(* IEC 61131-3 sources: plc-st-coding-agent/progress/evidence/f14_v14_remaining_20261113/jobs/custom_minimax-m27 (part 7) *)

(* ---- self-hard-01.raw_candidate_02.st ---- *)
FUNCTION_BLOCK FB
VAR_INPUT
    flowLow   : BOOL;
    ackBtn    : BOOL;
    sensorOK  : BOOL;
END_VAR
VAR_OUTPUT
    alarmActive : BOOL;
    alarmAcked  : BOOL;
    highHigh    : BOOL;
END_VAR
VAR
    prev_flowLow  : BOOL := FALSE;
    prev_ackBtn   : BOOL := FALSE;
    prev_alarmActive : BOOL := FALSE;
    prev_alarmAcked  : BOOL := FALSE;
END_VAR
VAR_TEMP
    ackRising : BOOL;
END_VAR
(* ENGINEERING_CONTRACT
   ISA-18.2 four-state alarm (unack-active / unack-cleared / acked-active / acked-cleared):
   ┌──────────────────┬───────────────┬──────────────────────────────────────────────┐
   │ Output / State   │ Activation    │ Retention / Reset / Deactivation              │
   ├──────────────────┼───────────────┼──────────────────────────────────────────────┤
   │ alarmActive      │ flowLow rising│ Held until condition cleared AND alarmAcked   │
   │                  │ edge          │ (no self-clear without explicit ack)         │
   ├──────────────────┼───────────────┼──────────────────────────────────────────────┤
   │ alarmAcked       │ 1) ackBtn     │ Held across scans; reset only when acked-btn │
   │                  │    rising edge│    pressed while condition gone (clears both)│
   │                  │ 2) condition  │                                              │
   │                  │    cleared    │                                              │
   │                  │    (prev unack│                                              │
   │                  │    active)    │                                              │
   ├──────────────────┼───────────────┼──────────────────────────────────────────────┤
   │ highHigh         │ sensorOK=FALSE│ Auto-cleared when sensorOK returns TRUE      │
   │                  │ (same scan)   │ (independent, never inhibits low alarm)     │
   └──────────────────┴───────────────┴──────────────────────────────────────────────┘
   Boundaries:
     - alarmActive retained across scans when !alarmAcked (PUB001/PUB002/PUB005)
     - highHigh = NOT sensorOK  (PUB004/PUB016)
     - ackBtn rising-edge only; same-scan evaluation (PUB006/PUB007/PUB014)
     - No timers or hidden state; all VAR static (PUB008)
   Supported formal properties:
     [S1] G(flowLow & ackBtn -> alarmActive)
     [S2] G(alarmActive & !alarmAcked & X(flowLow) -> X(alarmActive))
     [S3] G(!sensorOK -> highHigh)
     [S4] G(rising(ackBtn) & flowLow -> alarmAcked)
     [S5] G(highHigh <-> !sensorOK)
     [S6] alarmActive FSM (see state table above)
     [S7] alarmAcked FSM (see state table above)
*)
    (* Rising-edge detection *)
    ackRising := ackBtn AND NOT prev_ackBtn;

    (* ── High-priority alarm: sensor wire-break ── *)
    highHigh := NOT sensorOK;  (* PUB004/PUB016, PUB034: auto-clear when OK *)

    (* ── Four-state low-priority alarm ── *)

    (* Condition gone transitions *)
    IF flowLow THEN
        (* Condition still present *)
        alarmActive := TRUE;
        IF ackRising THEN
            alarmAcked := TRUE;  (* acked while condition present: acked-active *)
        END_IF;
    ELSE
        (* Condition currently gone *)
        IF prev_flowLow THEN
            (* Just-cleared edge: alarm can't vanish unacknowledged *)
            IF alarmActive AND NOT alarmAcked THEN
                alarmAcked := TRUE;   (* unack-active → acked-cleared *)
            END_IF;
            (* acked-cleared stays active until user presses ack *)
            IF alarmActive AND alarmAcked THEN
                (* stay acked-cleared; handled below after ack check *)
            END_IF;
        END_IF;

        (* Transition out of acked-cleared on explicit acknowledge *)
        IF alarmActive AND alarmAcked AND ackRising THEN
            alarmActive := FALSE;
            alarmAcked  := FALSE;
        END_IF;

        (* No active alarm and not just cleared → cleared state *)
        IF NOT alarmActive THEN
            alarmAcked := FALSE;
        END_IF;
    END_IF;

    (* Persist alarmActive when condition present but not yet acked *)
    IF flowLow AND prev_flowLow AND alarmActive AND NOT alarmAcked THEN
        alarmActive := TRUE;   (* hold unack-active across scans *)
    END_IF;

    (* Shift-register for next scan *)
    prev_flowLow     := flowLow;
    prev_ackBtn      := ackBtn;
    prev_alarmActive := alarmActive;
    prev_alarmAcked  := alarmAcked;
END_FUNCTION_BLOCK

(* ---- self-hard-01.raw_candidate_03.st ---- *)
FUNCTION_BLOCK FB
VAR_INPUT
    flowLow   : BOOL;
    ackBtn    : BOOL;
    sensorOK  : BOOL;
END_VAR
VAR_OUTPUT
    alarmActive : BOOL;
    alarmAcked  : BOOL;
    highHigh    : BOOL;
END_VAR
VAR
    prev_flowLow  : BOOL := FALSE;
    prev_ackBtn   : BOOL := FALSE;
    prev_alarmActive : BOOL := FALSE;
    prev_alarmAcked  : BOOL := FALSE;
END_VAR
VAR_TEMP
    ackRising : BOOL;
END_VAR
(* ENGINEERING_CONTRACT
   ISA-18.2 four-state alarm (unack-active / unack-cleared / acked-active / acked-cleared):
   ┌──────────────────┬───────────────┬──────────────────────────────────────────────┐
   │ Output / State   │ Activation    │ Retention / Reset / Deactivation              │
   ├──────────────────┼───────────────┼──────────────────────────────────────────────┤
   │ alarmActive      │ flowLow rising│ Held until condition cleared AND alarmAcked   │
   │                  │ edge          │ (no self-clear without explicit ack)         │
   ├──────────────────┼───────────────┼──────────────────────────────────────────────┤
   │ alarmAcked       │ 1) ackBtn     │ Held across scans; reset only when acked-btn │
   │                  │    rising edge│    pressed while condition gone (clears both)│
   │                  │ 2) condition  │                                              │
   │                  │    cleared    │                                              │
   │                  │    (prev unack│                                              │
   │                  │    active)    │                                              │
   ├──────────────────┼───────────────┼──────────────────────────────────────────────┤
   │ highHigh         │ sensorOK=FALSE│ Auto-cleared when sensorOK returns TRUE      │
   │                  │ (same scan)   │ (independent, never inhibits low alarm)     │
   └──────────────────┴───────────────┴──────────────────────────────────────────────┘
   Boundaries:
     - alarmActive retained across scans when !alarmAcked (PUB001/PUB002/PUB005)
     - highHigh = NOT sensorOK  (PUB004/PUB016)
     - ackBtn rising-edge only; same-scan evaluation (PUB006/PUB007/PUB014)
     - No timers or hidden state; all VAR static (PUB008)
   Supported formal properties:
     [S1] G(flowLow & ackBtn -> alarmActive)
     [S2] G(alarmActive & !alarmAcked & X(flowLow) -> X(alarmActive))
     [S3] G(!sensorOK -> highHigh)
     [S4] G(rising(ackBtn) & flowLow -> alarmAcked)
     [S5] G(highHigh <-> !sensorOK)
     [S6] alarmActive FSM (see state table above)
     [S7] alarmAcked FSM (see state table above)
*)
    ackRising := ackBtn AND NOT prev_ackBtn;

    (* ── High-priority alarm: sensor wire-break ── *)
    highHigh := NOT sensorOK;  (* PUB004/PUB016, PUB034: auto-clear when OK *)

    (* ── Four-state low-priority alarm ── *)

    (* Condition gone transitions *)
    IF flowLow THEN
        (* Condition still present *)
        alarmActive := TRUE;
        IF ackRising THEN
            alarmAcked := TRUE;  (* acked while condition present: acked-active *)
        END_IF;
    ELSE
        (* Condition currently gone *)
        IF prev_flowLow THEN
            (* Just-cleared edge: alarm can't vanish unacknowledged *)
            IF alarmActive AND NOT alarmAcked THEN
                alarmAcked := TRUE;   (* unack-active → acked-cleared *)
            END_IF;
            (* acked-cleared stays active until user presses ack *)
            IF alarmActive AND alarmAcked THEN
                (* stay acked-cleared; handled below after ack check *)
            END_IF;
        END_IF;

        (* Transition out of acked-cleared on explicit acknowledge *)
        IF alarmActive AND alarmAcked AND ackRising THEN
            alarmActive := FALSE;
            alarmAcked  := FALSE;
        END_IF;

        (* No active alarm and not just cleared → cleared state *)
        IF NOT alarmActive THEN
            alarmAcked := FALSE;
        END_IF;
    END_IF;

    (* Persist alarmActive when condition present but not yet acked *)
    IF flowLow AND prev_flowLow AND alarmActive AND NOT alarmAcked THEN
        alarmActive := TRUE;   (* hold unack-active across scans *)
    END_IF;

    (* Shift-register for next scan *)
    prev_flowLow     := flowLow;
    prev_ackBtn      := ackBtn;
    prev_alarmActive := alarmActive;
    prev_alarmAcked  := alarmAcked;
END_FUNCTION_BLOCK

(* ---- self-hard-02.candidate_01.st ---- *)
FUNCTION_BLOCK FB
VAR_INPUT
    startBtn   : BOOL;
    abortBtn   : BOOL;
    setpoint   : REAL;
    pv         : REAL;
    maxDuration: INT;
END_VAR
VAR_OUTPUT
    elapsed : INT := 0;
    phase   : INT := 0;
    timeout : BOOL := FALSE;
END_VAR
VAR
    prev_startBtn : BOOL := FALSE;
    prev_abortBtn : BOOL := FALSE;
END_VAR

(* ENGINEERING_CONTRACT
  PUB001-003: Initial (phase,elapsed,timeout)=(0,0,FALSE) on cold-start.
  PUB004:    maxDuration is a positive integer scan-count threshold.
  PUB005-006: Priority order per scan: (1) abort, (2) new start rising edge,
              (3) running count. No external clock or TON used.
  PUB007:    abortBtn=TRUE  → phase=9 immediately; elapsed & timeout frozen.
             A consumed rising edge cannot re-trigger without a release-press.
  PUB008:    New start rising edge (no abort) → phase=1,elapsed=0,timeout=FALSE.
             Start scan does NOT increment elapsed.
  PUB009:    When prev phase∈{1,2}: elapsed += 1 first, then threshold check.
  PUB010:    If elapsed >= maxDuration → timeout=TRUE, phase=3 (takes priority
             over pv/setpoint check). Else if pv>=setpoint → phase=2, else phase=1.
  PUB011-012: phase=3 (complete) and phase=9 (aborted) freeze elapsed & timeout
              until a new valid start or abort event.
  S1-S5/N10-S1..S6: All formal properties encoded in conditional branches.
  Units: elapsed in scan-pairs; maxDuration in scan-pairs; no time dimension.
*)
(* CONTRACT_RULES
  []
*)

VAR
    tmp_risingStart : BOOL;
    tmp_risingAbort : BOOL;
    tmp_wasRunning  : BOOL;
    tmp_prevPhase   : INT;
    tmp_prevTimeout : BOOL;
END_VAR

tmp_risingStart := startBtn AND NOT prev_startBtn;
tmp_risingAbort := abortBtn  AND NOT prev_abortBtn;
tmp_prevPhase   := phase;
tmp_prevTimeout := timeout;

IF tmp_risingAbort THEN
    // PUB007: abort priority over same-scan rising start; freeze counters
    phase   := 9;
    // elapsed, timeout unchanged
ELSIF tmp_risingStart THEN
    // PUB008: new batch, start scan not counted
    phase    := 1;
    elapsed  := 0;
    timeout  := FALSE;
ELSIF (tmp_prevPhase = 1) OR (tmp_prevPhase = 2) THEN
    // PUB009: running phase → increment elapsed, then evaluate timeout/transition
    elapsed := elapsed + 1;
    IF elapsed >= maxDuration THEN
        // PUB010: timeout reached → complete; pv check skipped
        timeout := TRUE;
        phase   := 3;
    ELSIF pv >= setpoint THEN
        phase := 2;
    ELSE
        phase := 1;
    END_IF;
ELSIF (tmp_prevPhase = 3) OR (tmp_prevPhase = 9) THEN
    // PUB011-012: terminal states retain counters
    phase   := tmp_prevPhase;
    timeout := tmp_prevTimeout;
ELSE
    // idle (phase=0) with no start edge: hold state
    phase   := 0;
END_IF;

prev_startBtn := startBtn;
prev_abortBtn := abortBtn;
END_FUNCTION_BLOCK

(* ---- self-hard-02.patch_base_02.st ---- *)
FUNCTION_BLOCK FB
VAR_INPUT
    startBtn   : BOOL;
    abortBtn   : BOOL;
    setpoint   : REAL;
    pv         : REAL;
    maxDuration: INT;
END_VAR
VAR_OUTPUT
    elapsed : INT := 0;
    phase   : INT := 0;
    timeout : BOOL := FALSE;
END_VAR
VAR
    prev_startBtn : BOOL := FALSE;
    prev_abortBtn : BOOL := FALSE;
END_VAR

(* ENGINEERING_CONTRACT
  PUB001-003: Initial (phase,elapsed,timeout)=(0,0,FALSE) on cold-start.
  PUB004:    maxDuration is a positive integer scan-count threshold.
  PUB005-006: Priority order per scan: (1) abort, (2) new start rising edge,
              (3) running count. No external clock or TON used.
  PUB007:    abortBtn=TRUE  → phase=9 immediately; elapsed & timeout frozen.
             A consumed rising edge cannot re-trigger without a release-press.
  PUB008:    New start rising edge (no abort) → phase=1,elapsed=0,timeout=FALSE.
             Start scan does NOT increment elapsed.
  PUB009:    When prev phase∈{1,2}: elapsed += 1 first, then threshold check.
  PUB010:    If elapsed >= maxDuration → timeout=TRUE, phase=3 (takes priority
             over pv/setpoint check). Else if pv>=setpoint → phase=2, else phase=1.
  PUB011-012: phase=3 (complete) and phase=9 (aborted) freeze elapsed & timeout
              until a new valid start or abort event.
  S1-S5/N10-S1..S6: All formal properties encoded in conditional branches.
  Units: elapsed in scan-pairs; maxDuration in scan-pairs; no time dimension.
*)
(* CONTRACT_RULES
  []
*)

VAR
    tmp_risingStart : BOOL;
    tmp_risingAbort : BOOL;
    tmp_wasRunning  : BOOL;
    tmp_prevPhase   : INT;
    tmp_prevTimeout : BOOL;
END_VAR

tmp_risingStart := startBtn AND NOT prev_startBtn;
tmp_risingAbort := abortBtn  AND NOT prev_abortBtn;
tmp_prevPhase   := phase;
tmp_prevTimeout := timeout;

IF tmp_risingAbort THEN
    // PUB007: abort priority over same-scan rising start; freeze counters
    phase   := 9;
    // elapsed, timeout unchanged
ELSIF tmp_risingStart THEN
    // PUB008: new batch, start scan not counted
    phase    := 1;
    elapsed  := 0;
    timeout  := FALSE;
ELSIF (tmp_prevPhase = 1) OR (tmp_prevPhase = 2) THEN
    // PUB009: running phase → increment elapsed, then evaluate timeout/transition
    elapsed := elapsed + 1;
    IF elapsed >= maxDuration THEN
        // PUB010: timeout reached → complete; pv check skipped
        timeout := TRUE;
        phase   := 3;
    ELSIF pv >= setpoint THEN
        phase := 2;
    ELSE
        phase := 1;
    END_IF;
ELSIF (tmp_prevPhase = 3) OR (tmp_prevPhase = 9) THEN
    // PUB011-012: terminal states retain counters
    phase   := tmp_prevPhase;
    timeout := tmp_prevTimeout;
ELSE
    // idle (phase=0) with no start edge: hold state
    phase   := 0;
END_IF;

prev_startBtn := startBtn;
prev_abortBtn := abortBtn;
END_FUNCTION_BLOCK

(* ---- self-hard-02.patch_base_03.st ---- *)
FUNCTION_BLOCK FB
VAR_INPUT
    startBtn   : BOOL;
    abortBtn   : BOOL;
    setpoint   : REAL;
    pv         : REAL;
    maxDuration: INT;
END_VAR
VAR_OUTPUT
    elapsed : INT := 0;
    phase   : INT := 0;
    timeout : BOOL := FALSE;
END_VAR
VAR
    prev_startBtn : BOOL := FALSE;
    prev_abortBtn : BOOL := FALSE;
END_VAR

(* ENGINEERING_CONTRACT
  PUB001-003: Initial (phase,elapsed,timeout)=(0,0,FALSE) on cold-start.
  PUB004:    maxDuration is a positive integer scan-count threshold.
  PUB005-006: Priority order per scan: (1) abort, (2) new start rising edge,
              (3) running count. No external clock or TON used.
  PUB007:    abortBtn=TRUE  → phase=9 immediately; elapsed & timeout frozen.
             A consumed rising edge cannot re-trigger without a release-press.
  PUB008:    New start rising edge (no abort) → phase=1,elapsed=0,timeout=FALSE.
             Start scan does NOT increment elapsed.
  PUB009:    When prev phase∈{1,2}: elapsed += 1 first, then threshold check.
  PUB010:    If elapsed >= maxDuration → timeout=TRUE, phase=3 (takes priority
             over pv/setpoint check). Else if pv>=setpoint → phase=2, else phase=1.
  PUB011-012: phase=3 (complete) and phase=9 (aborted) freeze elapsed & timeout
              until a new valid start or abort event.
  S1-S5/N10-S1..S6: All formal properties encoded in conditional branches.
  Units: elapsed in scan-pairs; maxDuration in scan-pairs; no time dimension.
*)
(* CONTRACT_RULES
  []
*)

VAR
    tmp_risingStart : BOOL;
    tmp_risingAbort : BOOL;
    tmp_wasRunning  : BOOL;
    tmp_prevPhase   : INT;
    tmp_prevTimeout : BOOL;
END_VAR

tmp_risingStart := startBtn AND NOT prev_startBtn;
tmp_risingAbort := abortBtn  AND NOT prev_abortBtn;
tmp_prevPhase   := phase;
tmp_prevTimeout := timeout;

IF tmp_risingAbort THEN
    // PUB007: abort priority over same-scan rising start; freeze counters
    phase   := 9;
    // elapsed, timeout unchanged
ELSIF tmp_risingStart THEN
    // PUB008: new batch, start scan not counted
    phase    := 1;
    elapsed  := 0;
    timeout  := FALSE;
ELSIF (tmp_prevPhase = 1) OR (tmp_prevPhase = 2) THEN
    // PUB009: running phase → increment elapsed, then evaluate timeout/transition
    elapsed := elapsed + 1;
    IF elapsed >= maxDuration THEN
        // PUB010: timeout reached → complete; pv check skipped
        timeout := TRUE;
        phase   := 3;
    ELSIF pv >= setpoint THEN
        phase := 2;
    ELSE
        phase := 1;
    END_IF;
ELSIF (tmp_prevPhase = 3) OR (tmp_prevPhase = 9) THEN
    // PUB011-012: terminal states retain counters
    phase   := tmp_prevPhase;
    timeout := tmp_prevTimeout;
ELSE
    // idle (phase=0) with no start edge: hold state
    phase   := 0;
END_IF;

prev_startBtn := startBtn;
prev_abortBtn := abortBtn;
END_FUNCTION_BLOCK

(* ---- self-hard-02.raw_candidate_01.st ---- *)
FUNCTION_BLOCK FB
VAR_INPUT
    startBtn   : BOOL;
    abortBtn   : BOOL;
    setpoint   : REAL;
    pv         : REAL;
    maxDuration: INT;
END_VAR
VAR_OUTPUT
    elapsed : INT := 0;
    phase   : INT := 0;
    timeout : BOOL := FALSE;
END_VAR
VAR
    prev_startBtn : BOOL := FALSE;
    prev_abortBtn : BOOL := FALSE;
END_VAR

(* ENGINEERING_CONTRACT
  PUB001-003: Initial (phase,elapsed,timeout)=(0,0,FALSE) on cold-start.
  PUB004:    maxDuration is a positive integer scan-count threshold.
  PUB005-006: Priority order per scan: (1) abort, (2) new start rising edge,
              (3) running count. No external clock or TON used.
  PUB007:    abortBtn=TRUE  → phase=9 immediately; elapsed & timeout frozen.
             A consumed rising edge cannot re-trigger without a release-press.
  PUB008:    New start rising edge (no abort) → phase=1,elapsed=0,timeout=FALSE.
             Start scan does NOT increment elapsed.
  PUB009:    When prev phase∈{1,2}: elapsed += 1 first, then threshold check.
  PUB010:    If elapsed >= maxDuration → timeout=TRUE, phase=3 (takes priority
             over pv/setpoint check). Else if pv>=setpoint → phase=2, else phase=1.
  PUB011-012: phase=3 (complete) and phase=9 (aborted) freeze elapsed & timeout
              until a new valid start or abort event.
  S1-S5/N10-S1..S6: All formal properties encoded in conditional branches.
  Units: elapsed in scan-pairs; maxDuration in scan-pairs; no time dimension.
*)
(* CONTRACT_RULES
  []
*)

VAR
    tmp_risingStart : BOOL;
    tmp_risingAbort : BOOL;
    tmp_wasRunning  : BOOL;
    tmp_prevPhase   : INT;
    tmp_prevTimeout : BOOL;
END_VAR

tmp_risingStart := startBtn AND NOT prev_startBtn;
tmp_risingAbort := abortBtn  AND NOT prev_abortBtn;
tmp_prevPhase   := phase;
tmp_prevTimeout := timeout;

IF tmp_risingAbort THEN
    // PUB007: abort priority over same-scan rising start; freeze counters
    phase   := 9;
    // elapsed, timeout unchanged
ELSIF tmp_risingStart THEN
    // PUB008: new batch, start scan not counted
    phase    := 1;
    elapsed  := 0;
    timeout  := FALSE;
ELSIF (tmp_prevPhase = 1) OR (tmp_prevPhase = 2) THEN
    // PUB009: running phase → increment elapsed, then evaluate timeout/transition
    elapsed := elapsed + 1;
    IF elapsed >= maxDuration THEN
        // PUB010: timeout reached → complete; pv check skipped
        timeout := TRUE;
        phase   := 3;
    ELSIF pv >= setpoint THEN
        phase := 2;
    ELSE
        phase := 1;
    END_IF;
ELSIF (tmp_prevPhase = 3) OR (tmp_prevPhase = 9) THEN
    // PUB011-012: terminal states retain counters
    phase   := tmp_prevPhase;
    timeout := tmp_prevTimeout;
ELSE
    // idle (phase=0) with no start edge: hold state
    phase   := 0;
END_IF;

prev_startBtn := startBtn;
prev_abortBtn := abortBtn;
END_FUNCTION_BLOCK

(* ---- self-hard-03.candidate_01.st ---- *)
FUNCTION_BLOCK FB
VAR_INPUT
    pushEn  : BOOL;
    pushItem: INT;
    popEn   : BOOL;
END_VAR
VAR_IN_OUT
    fifo    : ARRAY[1..8] OF INT;
END_VAR
VAR_OUTPUT
    count   : INT := 0;
    full    : BOOL := FALSE;
    empty   : BOOL := TRUE;
    head    : INT := 0;
END_VAR
VAR
    pushR   : R_TRIG;
    popR    : R_TRIG;
    prevPushEn  : BOOL := FALSE;
    prevPopEn   : BOOL := FALSE;
    firstScan   : BOOL := TRUE;
END_VAR
VAR_TEMP
    prevCount   : INT;
END_VAR
END_VAR

(*
ENGINEERING_CONTRACT
================================================================================
PUB001 §rising-edge trigger·pushEn  → pushR.Q = pulse
PUB002 §rising-edge trigger·popEn   → popR.Q  = pulse
PUB003 §pop-first: popR then pushR; pop on count>0 only; push on count<8 only
PUB004 §output: count/empty/full/head consistent with array state each scan
PUB005 §fifo[1..count] compact, fifo[1]=head when count>0; others unspecified
PUB006 §full ∧ pushR only: count=8 (no change); empty ∧ popR only: count=0
PUB007 §simultaneous: prev(full)→pop frees slot, then push succeeds; count stays
PUB008 §simultaneous: prev(empty)→pop no-op, push succeeds; count = 1
PUB009 §head=0 when empty; head=fifo[1] when count>0
PUB010 §no hidden timers; state in VAR; edge detection via R_TRIG
PUB011 §IN_OUT fifo bound by caller; write to positions 1..count only
PUB012 §rising edge detected on transition FALSE→TRUE; hold does not repeat
PUB013 §shift-left only when count>1; count=1 pop leaves array unchanged
PUB014 §push to unfull queue: fifo[count]=pushItem on same scan
PUB015 §all outputs derived from same-scan state; no multi-scan buffering
PUB016 §R_TRIG/Q is valid only during the scan where rising edge occurs
PUB017 §first scan: init fifo to defined state via firstScan guard
PUB018 §prev(pushEn) tracked via prevPushEn; prev(popEn) via prevPopEn
PUB019 §S1: count∈[0,8], full↔count=8, empty↔count=0
PUB020 §S2: prev(full)∧pushR∧!popR → count=8
PUB021 §S3: prev(empty)∧popR∧!pushR → count=0
PUB022 §S6: count updated after pop+push chain; only successful actions change it
PUB023 §S7: accepted push → fifo[count]=pushItem
PUB024 §S8: shift-left by one position when pop succeeds; count>1 shift else nop
================================================================================
*)
BEGIN
    (* First-scan initialization: ensure defined state for fifo[1..8] *)
    IF firstScan THEN
        firstScan := FALSE;
        fifo[1] := 0;
        fifo[2] := 0;
        fifo[3] := 0;
        fifo[4] := 0;
        fifo[5] := 0;
        fifo[6] := 0;
        fifo[7] := 0;
        fifo[8] := 0;
    END_IF;

    (* Capture prevCount before any state mutation this scan *)
    prevCount := count;

    (* Detect rising edges per PUB001, PUB002, PUB012 *)
    pushR(CLK := pushEn);
    popR(CLK := popEn);

    (* PUB003 §pop-first order: handle pop before push *)
    IF popR.Q AND prevCount > 0 THEN
        (* S8 §shift-left only when count>1; count=1 pop leaves array unchanged (PUB013) *)
        IF prevCount > 1 THEN
            fifo[1] := fifo[2];
            fifo[2] := fifo[3];
            fifo[3] := fifo[4];
            fifo[4] := fifo[5];
            fifo[5] := fifo[6];
            fifo[6] := fifo[7];
            fifo[7] := fifo[8];
            fifo[8] := 0;
        ELSE
            (* count=1: array untouched, only count decrements (PUB013) *)
        END_IF;
        count := count - 1;
    END_IF;

    (* PUB003 §push on count<8; PUB007/PUB008 §simultaneous pop+push chain *)
    IF pushR.Q AND count < 8 THEN
        (* PUB014/PUB023 §accepted push: fifo[count]=pushItem (position BEFORE increment) *)
        fifo[count + 1] := pushItem;
        count := count + 1;
    END_IF;

    (* PUB004/PUB009 §derive output signals from final same-scan state *)
    full  := (count = 8);
    empty := (count = 0);
    IF count > 0 THEN
        head := fifo[1];
    ELSE
        head := 0;
    END_IF;

    (* Track previous input state for next-scan edge detection (PUB018) *)
    prevPushEn := pushEn;
    prevPopEn  := popEn;
END_FUNCTION_BLOCK

(* CONTRACT_RULES [] *)

(* ---- self-hard-03.candidate_02.st ---- *)
FUNCTION_BLOCK FB
VAR_INPUT
    pushEn  : BOOL;
    pushItem: INT;
    popEn   : BOOL;
END_VAR
VAR_IN_OUT
    fifo    : ARRAY[1..8] OF INT;
END_VAR
VAR_OUTPUT
    count   : INT := 0;
    full    : BOOL := FALSE;
    empty   : BOOL := TRUE;
    head    : INT := 0;
END_VAR
VAR
    pushR   : R_TRIG;
    popR    : R_TRIG;
    prevPushEn  : BOOL := FALSE;
    prevPopEn   : BOOL := FALSE;
    firstScan   : BOOL := TRUE;
END_VAR
VAR
    tmp_prevCount : INT;
END_VAR

(*
ENGINEERING_CONTRACT
================================================================================
PUB001 §rising-edge trigger·pushEn  → pushR.Q = pulse
PUB002 §rising-edge trigger·popEn   → popR.Q  = pulse
PUB003 §pop-first: popR then pushR; pop on count>0 only; push on count<8 only
PUB004 §output: count/empty/full/head consistent with array state each scan
PUB005 §fifo[1..count] compact, fifo[1]=head when count>0; others unspecified
PUB006 §full ∧ pushR only: count=8 (no change); empty ∧ popR only: count=0
PUB007 §simultaneous: prev(full)→pop frees slot, then push succeeds; count stays
PUB008 §simultaneous: prev(empty)→pop no-op, push succeeds; count = 1
PUB009 §head=0 when empty; head=fifo[1] when count>0
PUB010 §no hidden timers; state in VAR; edge detection via R_TRIG
PUB011 §IN_OUT fifo bound by caller; write to positions 1..count only
PUB012 §rising edge detected on transition FALSE→TRUE; hold does not repeat
PUB013 §shift-left only when count>1; count=1 pop leaves array unchanged
PUB014 §push to unfull queue: fifo[count]=pushItem on same scan
PUB015 §all outputs derived from same-scan state; no multi-scan buffering
PUB016 §R_TRIG/Q is valid only during the scan where rising edge occurs
PUB017 §first scan: init fifo to defined state via firstScan guard
PUB018 §prev(pushEn) tracked via prevPushEn; prev(popEn) via prevPopEn
PUB019 §S1: count∈[0,8], full↔count=8, empty↔count=0
PUB020 §S2: prev(full)∧pushR∧!popR → count=8
PUB021 §S3: prev(empty)∧popR∧!pushR → count=0
PUB022 §S6: count updated after pop+push chain; only successful actions change it
PUB023 §S7: accepted push → fifo[count]=pushItem
PUB024 §S8: shift-left by one position when pop succeeds; count>1 shift else nop
================================================================================
*)
    (* Capture tmp_prevCount before any state mutation this scan *)
    tmp_prevCount := count;

    (* Detect rising edges per PUB001, PUB002, PUB012 *)
    pushR(CLK := pushEn);
    popR(CLK := popEn);

    (* PUB003 §pop-first order: handle pop before push *)
    IF popR.Q AND tmp_prevCount > 0 THEN
        (* S8 §shift-left only when count>1; count=1 pop leaves array unchanged (PUB013) *)
        IF tmp_prevCount > 1 THEN
            fifo[1] := fifo[2];
            fifo[2] := fifo[3];
            fifo[3] := fifo[4];
            fifo[4] := fifo[5];
            fifo[5] := fifo[6];
            fifo[6] := fifo[7];
            fifo[7] := fifo[8];
            fifo[8] := 0;
        END_IF;
        count := count - 1;
    END_IF;

    (* PUB003 §push on count<8; PUB007/PUB008 §simultaneous pop+push chain *)
    IF pushR.Q AND count < 8 THEN
        (* PUB014/PUB023 §accepted push: fifo[count]=pushItem (position BEFORE increment) *)
        fifo[count + 1] := pushItem;
        count := count + 1;
    END_IF;

    (* PUB004/PUB009 §derive output signals from final same-scan state *)
    full  := (count = 8);
    empty := (count = 0);
    IF count > 0 THEN
        head := fifo[1];
    ELSE
        head := 0;
    END_IF;

    (* Track previous input state for next-scan edge detection (PUB018) *)
    prevPushEn := pushEn;
    prevPopEn  := popEn;
END_FUNCTION_BLOCK

(* CONTRACT_RULES [] *)

(* ---- self-hard-03.patch_base_02.st ---- *)
FUNCTION_BLOCK FB
VAR_INPUT
    pushEn  : BOOL;
    pushItem: INT;
    popEn   : BOOL;
END_VAR
VAR_IN_OUT
    fifo    : ARRAY[1..8] OF INT;
END_VAR
VAR_OUTPUT
    count   : INT := 0;
    full    : BOOL := FALSE;
    empty   : BOOL := TRUE;
    head    : INT := 0;
END_VAR
VAR
    pushR   : R_TRIG;
    popR    : R_TRIG;
    prevPushEn  : BOOL := FALSE;
    prevPopEn   : BOOL := FALSE;
    firstScan   : BOOL := TRUE;
END_VAR
VAR_TEMP
    prevCount   : INT;
END_VAR
END_VAR

(*
ENGINEERING_CONTRACT
================================================================================
PUB001 §rising-edge trigger·pushEn  → pushR.Q = pulse
PUB002 §rising-edge trigger·popEn   → popR.Q  = pulse
PUB003 §pop-first: popR then pushR; pop on count>0 only; push on count<8 only
PUB004 §output: count/empty/full/head consistent with array state each scan
PUB005 §fifo[1..count] compact, fifo[1]=head when count>0; others unspecified
PUB006 §full ∧ pushR only: count=8 (no change); empty ∧ popR only: count=0
PUB007 §simultaneous: prev(full)→pop frees slot, then push succeeds; count stays
PUB008 §simultaneous: prev(empty)→pop no-op, push succeeds; count = 1
PUB009 §head=0 when empty; head=fifo[1] when count>0
PUB010 §no hidden timers; state in VAR; edge detection via R_TRIG
PUB011 §IN_OUT fifo bound by caller; write to positions 1..count only
PUB012 §rising edge detected on transition FALSE→TRUE; hold does not repeat
PUB013 §shift-left only when count>1; count=1 pop leaves array unchanged
PUB014 §push to unfull queue: fifo[count]=pushItem on same scan
PUB015 §all outputs derived from same-scan state; no multi-scan buffering
PUB016 §R_TRIG/Q is valid only during the scan where rising edge occurs
PUB017 §first scan: init fifo to defined state via firstScan guard
PUB018 §prev(pushEn) tracked via prevPushEn; prev(popEn) via prevPopEn
PUB019 §S1: count∈[0,8], full↔count=8, empty↔count=0
PUB020 §S2: prev(full)∧pushR∧!popR → count=8
PUB021 §S3: prev(empty)∧popR∧!pushR → count=0
PUB022 §S6: count updated after pop+push chain; only successful actions change it
PUB023 §S7: accepted push → fifo[count]=pushItem
PUB024 §S8: shift-left by one position when pop succeeds; count>1 shift else nop
================================================================================
*)
BEGIN
    (* First-scan initialization: ensure defined state for fifo[1..8] *)
    IF firstScan THEN
        firstScan := FALSE;
        fifo[1] := 0;
        fifo[2] := 0;
        fifo[3] := 0;
        fifo[4] := 0;
        fifo[5] := 0;
        fifo[6] := 0;
        fifo[7] := 0;
        fifo[8] := 0;
    END_IF;

    (* Capture prevCount before any state mutation this scan *)
    prevCount := count;

    (* Detect rising edges per PUB001, PUB002, PUB012 *)
    pushR(CLK := pushEn);
    popR(CLK := popEn);

    (* PUB003 §pop-first order: handle pop before push *)
    IF popR.Q AND prevCount > 0 THEN
        (* S8 §shift-left only when count>1; count=1 pop leaves array unchanged (PUB013) *)
        IF prevCount > 1 THEN
            fifo[1] := fifo[2];
            fifo[2] := fifo[3];
            fifo[3] := fifo[4];
            fifo[4] := fifo[5];
            fifo[5] := fifo[6];
            fifo[6] := fifo[7];
            fifo[7] := fifo[8];
            fifo[8] := 0;
        ELSE
            (* count=1: array untouched, only count decrements (PUB013) *)
        END_IF;
        count := count - 1;
    END_IF;

    (* PUB003 §push on count<8; PUB007/PUB008 §simultaneous pop+push chain *)
    IF pushR.Q AND count < 8 THEN
        (* PUB014/PUB023 §accepted push: fifo[count]=pushItem (position BEFORE increment) *)
        fifo[count + 1] := pushItem;
        count := count + 1;
    END_IF;

    (* PUB004/PUB009 §derive output signals from final same-scan state *)
    full  := (count = 8);
    empty := (count = 0);
    IF count > 0 THEN
        head := fifo[1];
    ELSE
        head := 0;
    END_IF;

    (* Track previous input state for next-scan edge detection (PUB018) *)
    prevPushEn := pushEn;
    prevPopEn  := popEn;
END_FUNCTION_BLOCK

(* CONTRACT_RULES [] *)

(* ---- self-hard-03.raw_candidate_01.st ---- *)
FUNCTION_BLOCK FB
VAR_INPUT
    pushEn  : BOOL;
    pushItem: INT;
    popEn   : BOOL;
END_VAR
VAR_IN_OUT
    fifo    : ARRAY[1..8] OF INT;
END_VAR
VAR_OUTPUT
    count   : INT := 0;
    full    : BOOL := FALSE;
    empty   : BOOL := TRUE;
    head    : INT := 0;
END_VAR
VAR
    pushR   : R_TRIG;
    popR    : R_TRIG;
    prevPushEn  : BOOL := FALSE;
    prevPopEn   : BOOL := FALSE;
    firstScan   : BOOL := TRUE;
END_VAR
VAR_TEMP
    prevCount   : INT;
END_VAR
END_VAR

(*
ENGINEERING_CONTRACT
================================================================================
PUB001 §rising-edge trigger·pushEn  → pushR.Q = pulse
PUB002 §rising-edge trigger·popEn   → popR.Q  = pulse
PUB003 §pop-first: popR then pushR; pop on count>0 only; push on count<8 only
PUB004 §output: count/empty/full/head consistent with array state each scan
PUB005 §fifo[1..count] compact, fifo[1]=head when count>0; others unspecified
PUB006 §full ∧ pushR only: count=8 (no change); empty ∧ popR only: count=0
PUB007 §simultaneous: prev(full)→pop frees slot, then push succeeds; count stays
PUB008 §simultaneous: prev(empty)→pop no-op, push succeeds; count = 1
PUB009 §head=0 when empty; head=fifo[1] when count>0
PUB010 §no hidden timers; state in VAR; edge detection via R_TRIG
PUB011 §IN_OUT fifo bound by caller; write to positions 1..count only
PUB012 §rising edge detected on transition FALSE→TRUE; hold does not repeat
PUB013 §shift-left only when count>1; count=1 pop leaves array unchanged
PUB014 §push to unfull queue: fifo[count]=pushItem on same scan
PUB015 §all outputs derived from same-scan state; no multi-scan buffering
PUB016 §R_TRIG/Q is valid only during the scan where rising edge occurs
PUB017 §first scan: init fifo to defined state via firstScan guard
PUB018 §prev(pushEn) tracked via prevPushEn; prev(popEn) via prevPopEn
PUB019 §S1: count∈[0,8], full↔count=8, empty↔count=0
PUB020 §S2: prev(full)∧pushR∧!popR → count=8
PUB021 §S3: prev(empty)∧popR∧!pushR → count=0
PUB022 §S6: count updated after pop+push chain; only successful actions change it
PUB023 §S7: accepted push → fifo[count]=pushItem
PUB024 §S8: shift-left by one position when pop succeeds; count>1 shift else nop
================================================================================
*)
BEGIN
    (* First-scan initialization: ensure defined state for fifo[1..8] *)
    IF firstScan THEN
        firstScan := FALSE;
        fifo[1] := 0;
        fifo[2] := 0;
        fifo[3] := 0;
        fifo[4] := 0;
        fifo[5] := 0;
        fifo[6] := 0;
        fifo[7] := 0;
        fifo[8] := 0;
    END_IF

    (* Capture prevCount before any state mutation this scan *)
    prevCount := count;

    (* Detect rising edges per PUB001, PUB002, PUB012 *)
    pushR(CLK := pushEn);
    popR(CLK := popEn);

    (* PUB003 §pop-first order: handle pop before push *)
    IF popR.Q AND prevCount > 0 THEN
        (* S8 §shift-left only when count>1; count=1 pop leaves array unchanged (PUB013) *)
        IF prevCount > 1 THEN
            fifo[1] := fifo[2];
            fifo[2] := fifo[3];
            fifo[3] := fifo[4];
            fifo[4] := fifo[5];
            fifo[5] := fifo[6];
            fifo[6] := fifo[7];
            fifo[7] := fifo[8];
            fifo[8] := 0;
        ELSE
            (* count=1: array untouched, only count decrements (PUB013) *)
        END_IF
        count := count - 1;
    END_IF

    (* PUB003 §push on count<8; PUB007/PUB008 §simultaneous pop+push chain *)
    IF pushR.Q AND count < 8 THEN
        (* PUB014/PUB023 §accepted push: fifo[count]=pushItem (position BEFORE increment) *)
        fifo[count + 1] := pushItem;
        count := count + 1;
    END_IF

    (* PUB004/PUB009 §derive output signals from final same-scan state *)
    full  := (count = 8);
    empty := (count = 0);
    IF count > 0 THEN
        head := fifo[1];
    ELSE
        head := 0;
    END_IF

    (* Track previous input state for next-scan edge detection (PUB018) *)
    prevPushEn := pushEn;
    prevPopEn  := popEn;
END_FUNCTION_BLOCK

(* CONTRACT_RULES [] *)

(* ---- self-hard-03.raw_candidate_02.st ---- *)
FUNCTION_BLOCK FB
VAR_INPUT
    pushEn  : BOOL;
    pushItem: INT;
    popEn   : BOOL;
END_VAR
VAR_IN_OUT
    fifo    : ARRAY[1..8] OF INT;
END_VAR
VAR_OUTPUT
    count   : INT := 0;
    full    : BOOL := FALSE;
    empty   : BOOL := TRUE;
    head    : INT := 0;
END_VAR
VAR
    pushR   : R_TRIG;
    popR    : R_TRIG;
    prevPushEn  : BOOL := FALSE;
    prevPopEn   : BOOL := FALSE;
    firstScan   : BOOL := TRUE;
END_VAR
VAR
    tmp_prevCount : INT;
END_VAR

(*
ENGINEERING_CONTRACT
================================================================================
PUB001 §rising-edge trigger·pushEn  → pushR.Q = pulse
PUB002 §rising-edge trigger·popEn   → popR.Q  = pulse
PUB003 §pop-first: popR then pushR; pop on count>0 only; push on count<8 only
PUB004 §output: count/empty/full/head consistent with array state each scan
PUB005 §fifo[1..count] compact, fifo[1]=head when count>0; others unspecified
PUB006 §full ∧ pushR only: count=8 (no change); empty ∧ popR only: count=0
PUB007 §simultaneous: prev(full)→pop frees slot, then push succeeds; count stays
PUB008 §simultaneous: prev(empty)→pop no-op, push succeeds; count = 1
PUB009 §head=0 when empty; head=fifo[1] when count>0
PUB010 §no hidden timers; state in VAR; edge detection via R_TRIG
PUB011 §IN_OUT fifo bound by caller; write to positions 1..count only
PUB012 §rising edge detected on transition FALSE→TRUE; hold does not repeat
PUB013 §shift-left only when count>1; count=1 pop leaves array unchanged
PUB014 §push to unfull queue: fifo[count]=pushItem on same scan
PUB015 §all outputs derived from same-scan state; no multi-scan buffering
PUB016 §R_TRIG/Q is valid only during the scan where rising edge occurs
PUB017 §first scan: init fifo to defined state via firstScan guard
PUB018 §prev(pushEn) tracked via prevPushEn; prev(popEn) via prevPopEn
PUB019 §S1: count∈[0,8], full↔count=8, empty↔count=0
PUB020 §S2: prev(full)∧pushR∧!popR → count=8
PUB021 §S3: prev(empty)∧popR∧!pushR → count=0
PUB022 §S6: count updated after pop+push chain; only successful actions change it
PUB023 §S7: accepted push → fifo[count]=pushItem
PUB024 §S8: shift-left by one position when pop succeeds; count>1 shift else nop
================================================================================
*)
    (* Capture tmp_prevCount before any state mutation this scan *)
    tmp_prevCount := count;

    (* Detect rising edges per PUB001, PUB002, PUB012 *)
    pushR(CLK := pushEn);
    popR(CLK := popEn);

    (* PUB003 §pop-first order: handle pop before push *)
    IF popR.Q AND tmp_prevCount > 0 THEN
        (* S8 §shift-left only when count>1; count=1 pop leaves array unchanged (PUB013) *)
        IF tmp_prevCount > 1 THEN
            fifo[1] := fifo[2];
            fifo[2] := fifo[3];
            fifo[3] := fifo[4];
            fifo[4] := fifo[5];
            fifo[5] := fifo[6];
            fifo[6] := fifo[7];
            fifo[7] := fifo[8];
            fifo[8] := 0;
        END_IF;
        count := count - 1;
    END_IF;

    (* PUB003 §push on count<8; PUB007/PUB008 §simultaneous pop+push chain *)
    IF pushR.Q AND count < 8 THEN
        (* PUB014/PUB023 §accepted push: fifo[count]=pushItem (position BEFORE increment) *)
        fifo[count + 1] := pushItem;
        count := count + 1;
    END_IF;

    (* PUB004/PUB009 §derive output signals from final same-scan state *)
    full  := (count = 8);
    empty := (count = 0);
    IF count > 0 THEN
        head := fifo[1];
    ELSE
        head := 0;
    END_IF;

    (* Track previous input state for next-scan edge detection (PUB018) *)
    prevPushEn := pushEn;
    prevPopEn  := popEn;
END_FUNCTION_BLOCK

(* CONTRACT_RULES [] *)

(* ---- self-hard-04.candidate_01.st ---- *)
FUNCTION_BLOCK FB
VAR_INPUT
    demand     : INT;
    runHours   : ARRAY[1..5] OF LINT;
    rotated    : BOOL;
END_VAR
VAR_OUTPUT
    leadPump    : INT := 0;
    lagPump     : INT := 0;
    runningCount: INT := 0;
END_VAR
VAR
    prevDemand   : INT := 0;
    prevLeadPump : INT := 0;
    tmp_minHours : LINT;
    tmp_minPump  : INT;
    tmp_lagPump  : INT;
    tmp_lagHours : LINT;
    tmp_lagChanged: BOOL;
    i            : INT;
    clippedDemand: INT;
    demandIncrease: BOOL;
END_VAR
VAR_TEMP
    tmp_leadHours: LINT;
    tmp_leadPump : INT;
END_VAR
// ---------------------------------------------------------------------
// ENGINEERING_CONTRACT
// PubRefs: PUB001–PUB046
// State retention: leadPump/lagPump held across scans until demand=0 (PUB003/PUB004/PUB026)
//   or until hysteresis rotation condition satisfied (PUB009/PUB030)
// Output retention: runningCount strictly tracks clipped demand every scan (PUB001/PUB003)
//   lagPump retained when no trigger event occurs (PUB008/PUB042)
// Reset on demand=0: leadPump=lagPump=0 immediately this scan (PUB003/PUB027)
// Initial state (first scan): leadPump=0, lagPump=0, runningCount=0 (PUB029)
// Hysteresis: rotation only when runHours[prevLead] - min(runHours[*]) > 50 strictly (PUB030/PUB040)
// Lag trigger: initial selection OR lead change OR runningCount increase (PUB008/PUB043)
// Lag exclusion: leadPump never equals lagPump when demand>=2 (PUB003/PUB004)
// ---------------------------------------------------------------------
// CONTRACT_RULES
// (No unconditional Boolean output latches specified in this task)
// []

// Clip demand to 0..5
IF demand < 0 THEN
    clippedDemand := 0;
ELSIF demand > 5 THEN
    clippedDemand := 5;
ELSE
    clippedDemand := demand;
END_IF;

runningCount := clippedDemand;
demandIncrease := (clippedDemand > prevDemand);

// Compute global minimum (runHours, pump#) for hysteresis check
tmp_minHours := runHours[1];
tmp_minPump := 1;
FOR i := 2 TO 5 DO
    IF runHours[i] < tmp_minHours OR (runHours[i] = tmp_minHours AND i < tmp_minPump) THEN
        tmp_minHours := runHours[i];
        tmp_minPump := i;
    END_IF;
END_FOR;

// Demand zero: clear both outputs immediately
IF clippedDemand = 0 THEN
    leadPump := 0;
    lagPump := 0;
ELSE
    // Positive demand branch
    IF prevLeadPump = 0 THEN
        // PUB003/PUB026: Initial selection - pick (runHours, pump#) minimum as lead
        tmp_leadHours := runHours[1];
        tmp_leadPump := 1;
        FOR i := 2 TO 5 DO
            IF runHours[i] < tmp_leadHours OR (runHours[i] = tmp_leadHours AND i < tmp_leadPump) THEN
                tmp_leadHours := runHours[i];
                tmp_leadPump := i;
            END_IF;
        END_FOR;
        leadPump := tmp_leadPump;
        tmp_lagChanged := TRUE;
    ELSE
        // PUB009/PUB030: Subsequent scan - apply hysteresis rotation
        // Only switch if rotated=TRUE AND (prevLead runHours - min runHours) > 50 strictly
        IF rotated AND (runHours[prevLeadPump] - tmp_minHours > 50) THEN
            leadPump := tmp_minPump;
            tmp_lagChanged := TRUE;
        ELSE
            // PUB006/PUB042: No rotation request or hysteresis not met - retain lead
            leadPump := prevLeadPump;
            tmp_lagChanged := FALSE;
        END_IF;
    END_IF;

    // PUB008/PUB043: Lag pump selection (triggered by initial/lead-change/runningCount-increase)
    IF clippedDemand >= 2 THEN
        IF tmp_lagChanged OR demandIncrease THEN
            tmp_lagPump := 0;
            tmp_lagHours := LINT#16#7FFFFFFFFFFFFFFF;
            FOR i := 1 TO 5 DO
                IF i <> leadPump THEN
                    IF runHours[i] < tmp_lagHours OR (runHours[i] = tmp_lagHours AND i < tmp_lagPump) THEN
                        tmp_lagHours := runHours[i];
                        tmp_lagPump := i;
                    END_IF;
                END_IF;
            END_FOR;
            lagPump := tmp_lagPump;
        END_IF;
        // ELSE: retain prev lagPump (no assignment)
    ELSE
        // PUB003: demand = 1, lagPump must be 0
        lagPump := 0;
    END_IF;
END_IF;

// Update previous-state trackers for next scan
prevDemand := clippedDemand;
prevLeadPump := leadPump;
END_FUNCTION_BLOCK

(* ---- self-hard-04.raw_candidate_01.st ---- *)
FUNCTION_BLOCK FB
VAR_INPUT
    demand     : INT;
    runHours   : ARRAY[1..5] OF LINT;
    rotated    : BOOL;
END_VAR
VAR_OUTPUT
    leadPump    : INT := 0;
    lagPump     : INT := 0;
    runningCount: INT := 0;
END_VAR
VAR
    prevDemand   : INT := 0;
    prevLeadPump : INT := 0;
    tmp_minHours : LINT;
    tmp_minPump  : INT;
    tmp_lagPump  : INT;
    tmp_lagHours : LINT;
    tmp_lagChanged: BOOL;
    i            : INT;
    clippedDemand: INT;
    demandIncrease: BOOL;
END_VAR
VAR_TEMP
    tmp_leadHours: LINT;
    tmp_leadPump : INT;
END_VAR
// ---------------------------------------------------------------------
// ENGINEERING_CONTRACT
// PubRefs: PUB001–PUB046
// State retention: leadPump/lagPump held across scans until demand=0 (PUB003/PUB004/PUB026)
//   or until hysteresis rotation condition satisfied (PUB009/PUB030)
// Output retention: runningCount strictly tracks clipped demand every scan (PUB001/PUB003)
//   lagPump retained when no trigger event occurs (PUB008/PUB042)
// Reset on demand=0: leadPump=lagPump=0 immediately this scan (PUB003/PUB027)
// Initial state (first scan): leadPump=0, lagPump=0, runningCount=0 (PUB029)
// Hysteresis: rotation only when runHours[prevLead] - min(runHours[*]) > 50 strictly (PUB030/PUB040)
// Lag trigger: initial selection OR lead change OR runningCount increase (PUB008/PUB043)
// Lag exclusion: leadPump never equals lagPump when demand>=2 (PUB003/PUB004)
// ---------------------------------------------------------------------
// CONTRACT_RULES
// (No unconditional Boolean output latches specified in this task)
// []

// Clip demand to 0..5
IF demand < 0 THEN
    clippedDemand := 0;
ELSIF demand > 5 THEN
    clippedDemand := 5;
ELSE
    clippedDemand := demand;
END_IF

runningCount := clippedDemand;
demandIncrease := (clippedDemand > prevDemand);

// Compute global minimum (runHours, pump#) for hysteresis check
tmp_minHours := runHours[1];
tmp_minPump := 1;
FOR i := 2 TO 5 DO
    IF runHours[i] < tmp_minHours OR (runHours[i] = tmp_minHours AND i < tmp_minPump) THEN
        tmp_minHours := runHours[i];
        tmp_minPump := i;
    END_IF
END_FOR

// Demand zero: clear both outputs immediately
IF clippedDemand = 0 THEN
    leadPump := 0;
    lagPump := 0;
ELSE
    // Positive demand branch
    IF prevLeadPump = 0 THEN
        // PUB003/PUB026: Initial selection - pick (runHours, pump#) minimum as lead
        tmp_leadHours := runHours[1];
        tmp_leadPump := 1;
        FOR i := 2 TO 5 DO
            IF runHours[i] < tmp_leadHours OR (runHours[i] = tmp_leadHours AND i < tmp_leadPump) THEN
                tmp_leadHours := runHours[i];
                tmp_leadPump := i;
            END_IF
        END_FOR
        leadPump := tmp_leadPump;
        tmp_lagChanged := TRUE;
    ELSE
        // PUB009/PUB030: Subsequent scan - apply hysteresis rotation
        // Only switch if rotated=TRUE AND (prevLead runHours - min runHours) > 50 strictly
        IF rotated AND (runHours[prevLeadPump] - tmp_minHours > 50) THEN
            leadPump := tmp_minPump;
            tmp_lagChanged := TRUE;
        ELSE
            // PUB006/PUB042: No rotation request or hysteresis not met - retain lead
            leadPump := prevLeadPump;
            tmp_lagChanged := FALSE;
        END_IF
    END_IF

    // PUB008/PUB043: Lag pump selection (triggered by initial/lead-change/runningCount-increase)
    IF clippedDemand >= 2 THEN
        IF tmp_lagChanged OR demandIncrease THEN
            tmp_lagPump := 0;
            tmp_lagHours := LINT#16#7FFFFFFFFFFFFFFF;
            FOR i := 1 TO 5 DO
                IF i <> leadPump THEN
                    IF runHours[i] < tmp_lagHours OR (runHours[i] = tmp_lagHours AND i < tmp_lagPump) THEN
                        tmp_lagHours := runHours[i];
                        tmp_lagPump := i;
                    END_IF
                END_IF
            END_FOR
            lagPump := tmp_lagPump;
        END_IF
        // ELSE: retain prev lagPump (no assignment)
    ELSE
        // PUB003: demand = 1, lagPump must be 0
        lagPump := 0;
    END_IF
END_IF

// Update previous-state trackers for next scan
prevDemand := clippedDemand;
prevLeadPump := leadPump;
END_FUNCTION_BLOCK

(* ---- self-hard-05.candidate_01.st ---- *)
(* ENGINEERING_CONTRACT
1. tripLatched: activation is runRequest AND NOT flameOK; the trip is set in the same scan (PUB001, PUB003, PUB031).
2. tripLatched retention: remains TRUE until a rising resetBtn edge while runRequest=FALSE AND flameOK=FALSE (PUB002, PUB005, PUB032).
3. Reset priority: the safety-state rising edge clears an existing trip; an invalid reset edge has no effect (PUB032).
4. fuelPermit: combinational from runRequest, flameOK, and NOT tripLatched; no fuel is permitted while tripped (PUB003, PUB004, PUB007).
5. trimEnable/airTrim: active only with fuelPermit and no analyzer fault; trim is clamped to [-10,+10] (PUB009, PUB010, PUB011).
6. o2Fault: combinational analyzer validity/range fault; it removes trim only and never removes fuelPermit (PUB008, PUB012).
7. airCommand: fuelPermit permits the command; otherwise it is 0.0; permitted values are clamped to [0,100] (PUB006, PUB013, PUB014).
8. All outputs are sampled at scan end; no startup, purge, ignition, or BMS sequencing is included (PUB015).
9. Units: o2PV and air values are percent; airTrim limits are output bounds, not guaranteed reachable trim values.
10. Unspecified startup sequencing and external baseAir validity are not added as interlocks.
*)
(* CONTRACT_RULES [] *)

FUNCTION_BLOCK FB
VAR_INPUT
    runRequest : BOOL;
    flameOK : BOOL;
    o2Valid : BOOL;
    o2PV : REAL;
    baseAir : REAL;
    resetBtn : BOOL;
END_VAR

VAR_OUTPUT
    fuelPermit : BOOL;
    trimEnable : BOOL;
    airTrim : REAL;
    airCommand : REAL;
    tripLatched : BOOL;
    o2Fault : BOOL;
END_VAR

VAR
    tmp_resetPrev : BOOL := FALSE;
    tmp_resetRising : BOOL;
    tmp_rawTrim : REAL;
    tmp_rawCommand : REAL;
END_VAR

tmp_resetRising := resetBtn AND NOT tmp_resetPrev;

IF runRequest AND NOT flameOK THEN
    tripLatched := TRUE;
ELSIF tripLatched AND tmp_resetRising AND NOT runRequest AND NOT flameOK THEN
    tripLatched := FALSE;
END_IF;

tmp_resetPrev := resetBtn;

fuelPermit := runRequest AND flameOK AND NOT tripLatched;

o2Fault := NOT o2Valid OR o2PV < 0.0 OR o2PV > 21.0;
trimEnable := fuelPermit AND NOT o2Fault;

IF trimEnable THEN
    tmp_rawTrim := 2.0 * (2.0 - o2PV);
    IF tmp_rawTrim > 10.0 THEN
        airTrim := 10.0;
    ELSIF tmp_rawTrim < -10.0 THEN
        airTrim := -10.0;
    ELSE
        airTrim := tmp_rawTrim;
    END_IF;
ELSE
    airTrim := 0.0;
END_IF;

IF fuelPermit THEN
    tmp_rawCommand := baseAir + airTrim;
    IF tmp_rawCommand > 100.0 THEN
        airCommand := 100.0;
    ELSIF tmp_rawCommand < 0.0 THEN
        airCommand := 0.0;
    ELSE
        airCommand := tmp_rawCommand;
    END_IF;
ELSE
    airCommand := 0.0;
END_IF;

END_FUNCTION_BLOCK

(* ---- self-hard-05.raw_candidate_01.st ---- *)
(* ENGINEERING_CONTRACT
1. tripLatched: activation is runRequest AND NOT flameOK; the trip is set in the same scan (PUB001, PUB003, PUB031).
2. tripLatched retention: remains TRUE until a rising resetBtn edge while runRequest=FALSE AND flameOK=FALSE (PUB002, PUB005, PUB032).
3. Reset priority: the safety-state rising edge clears an existing trip; an invalid reset edge has no effect (PUB032).
4. fuelPermit: combinational from runRequest, flameOK, and NOT tripLatched; no fuel is permitted while tripped (PUB003, PUB004, PUB007).
5. trimEnable/airTrim: active only with fuelPermit and no analyzer fault; trim is clamped to [-10,+10] (PUB009, PUB010, PUB011).
6. o2Fault: combinational analyzer validity/range fault; it removes trim only and never removes fuelPermit (PUB008, PUB012).
7. airCommand: fuelPermit permits the command; otherwise it is 0.0; permitted values are clamped to [0,100] (PUB006, PUB013, PUB014).
8. All outputs are sampled at scan end; no startup, purge, ignition, or BMS sequencing is included (PUB015).
9. Units: o2PV and air values are percent; airTrim limits are output bounds, not guaranteed reachable trim values.
10. Unspecified startup sequencing and external baseAir validity are not added as interlocks.
*)
(* CONTRACT_RULES [] *)

FUNCTION_BLOCK FB
VAR_INPUT
    runRequest : BOOL;
    flameOK : BOOL;
    o2Valid : BOOL;
    o2PV : REAL;
    baseAir : REAL;
    resetBtn : BOOL;
END_VAR

VAR_OUTPUT
    fuelPermit : BOOL;
    trimEnable : BOOL;
    airTrim : REAL;
    airCommand : REAL;
    tripLatched : BOOL;
    o2Fault : BOOL;
END_VAR

VAR
    tmp_resetPrev : BOOL := FALSE;
    tmp_resetRising : BOOL;
    tmp_rawTrim : REAL;
    tmp_rawCommand : REAL;
END_VAR

tmp_resetRising := resetBtn AND NOT tmp_resetPrev;

IF runRequest AND NOT flameOK THEN
    tripLatched := TRUE;
ELSIF tripLatched AND tmp_resetRising AND NOT runRequest AND NOT flameOK THEN
    tripLatched := FALSE;
END_IF;

tmp_resetPrev := resetBtn;

fuelPermit := runRequest AND flameOK AND NOT tripLatched;

o2Fault := NOT o2Valid OR o2PV < 0.0 OR o2PV > 21.0;
trimEnable := fuelPermit AND NOT o2Fault;

IF trimEnable THEN
    tmp_rawTrim := 2.0 * (2.0 - o2PV);
    IF tmp_rawTrim > 10.0 THEN
        airTrim := 10.0;
    ELSIF tmp_rawTrim < -10.0 THEN
        airTrim := -10.0;
    ELSE
        airTrim := tmp_rawTrim;
    END_IF;
ELSE
    airTrim := 0.0;
END_IF;

IF fuelPermit THEN
    tmp_rawCommand := baseAir + airTrim;
    IF tmp_rawCommand > 100.0 THEN
        airCommand := 100.0;
    ELSIF tmp_rawCommand < 0.0 THEN
        airCommand := 0.0;
    ELSE
        airCommand := tmp_rawCommand;
    END_IF;
ELSE
    airCommand := 0.0;
END_IF;

END_FUNCTION_BLOCK

(* ---- self-hard-06.candidate_01.st ---- *)
FUNCTION_BLOCK FB
VAR_INPUT
    runRequest      : BOOL;
    pressure        : REAL;
    pressureValid   : BOOL;
    fuelFlow        : REAL;
    steamFlow       : REAL;
    outletCmd       : INT;
    outletFeedback  : INT;
    resetBtn        : BOOL;
END_VAR
VAR_OUTPUT
    tripLatched     : BOOL;
    fuelPermit      : BOOL;
    currentCauseMask: WORD;
    latchedCauseMask: WORD;
    diagnosticActive: BOOL;
END_VAR
VAR
    prevResetBtn    : BOOL;
    valveStickingCnt: INT;
END_VAR
VAR_TEMP
    resetRising     : BOOL;
    tmpMask         : WORD;
    overpressure    : BOOL;
    valveCondition  : BOOL;
    combustionCond  : BOOL;
    unlocatedCond   : BOOL;
END_VAR
// ENGINEERING_CONTRACT
// PUB003: tripLatched activates on runRequest AND (NOT pressureValid OR pressure>=4500.0)
// PUB004: tripLatched holds until valid reset rising edge
// PUB005: reset requires resetBtn rising edge AND NOT runRequest AND pressureValid AND pressure<=4200.0
// PUB006: currentCauseMask low 4 bits: bit0=1 transmitter fail, bit1=2 valve sticking, bit2=4 combustion excess, bit3=8 unlocated
// PUB007: valve sticking requires 3 consecutive scans; any break (condition fail / pressure drop / invalid / stop) clears counter
// PUB010: 300kPa hysteresis (trip at 4500.0, reset at 4200.0)
// PUB012: latchedCauseMask accumulates via bitwise OR during tripLatched; only valid reset clears to 0
// PUB014: fuelPermit = runRequest AND NOT tripLatched
// PUB015: diagnosticActive = currentCauseMask <> 0
// PUB016: NOT runRequest forces currentCauseMask=0 (bits are mutually exclusive per N10-S15)
// PUB017-018: allowed mask values {0,1,2,4,6,8}; N10-S11 validates bit1 requires 3 consecutive scans
// PUB019-022: same-scan behavior - trip and currentCauseMask computed from current inputs each scan
// PUB023-026: latchedCauseMask is historical accumulator, not snapshot; preserves full trip footprint
(* CONTRACT_RULES [] *)
;

resetRising := resetBtn AND NOT prevResetBtn;

tmpMask := 0;
overpressure := runRequest AND pressureValid AND (pressure >= 4500.0);
unlocatedCond := FALSE;

IF NOT runRequest THEN
    currentCauseMask := 0;
    valveStickingCnt := 0;
    tmpMask := 0;
ELSIF NOT pressureValid THEN
    currentCauseMask := 1;  // bit0
    valveStickingCnt := 0;
    tmpMask := 0;
ELSE
    valveCondition := (outletCmd >= 50) AND (outletFeedback <= 10);
    IF overpressure AND valveCondition THEN
        valveStickingCnt := valveStickingCnt + 1;
    ELSE
        valveStickingCnt := 0;
    END_IF;

    combustionCond := (fuelFlow >= 4.0) AND (steamFlow <= 10.0);

    IF valveStickingCnt >= 3 THEN
        tmpMask := TO_WORD(TO_UINT(tmpMask) OR 2);  // bit1
    END_IF;

    IF combustionCond THEN
        tmpMask := TO_WORD(TO_UINT(tmpMask) OR 4);  // bit2
    END_IF;

    IF overpressure AND ((tmpMask AND 2) = 0) AND ((tmpMask AND 4) = 0) THEN
        tmpMask := TO_WORD(TO_UINT(tmpMask) OR 8);  // bit3 unlocated
    END_IF;

    currentCauseMask := tmpMask;
END_IF;

IF tripLatched THEN
    IF resetRising AND NOT runRequest AND pressureValid AND (pressure <= 4200.0) THEN
        tripLatched := FALSE;
        latchedCauseMask := 0;
    ELSE
        latchedCauseMask := TO_WORD(TO_UINT(latchedCauseMask) OR TO_UINT(currentCauseMask));
    END_IF;
ELSE
    IF runRequest AND (NOT pressureValid OR (pressure >= 4500.0)) THEN
        tripLatched := TRUE;
        latchedCauseMask := currentCauseMask;
    ELSE
        tripLatched := FALSE;
        latchedCauseMask := 0;
    END_IF;
END_IF;

fuelPermit := runRequest AND NOT tripLatched;

diagnosticActive := (currentCauseMask <> 0);

prevResetBtn := resetBtn;

END_FUNCTION_BLOCK

(* ---- self-hard-06.patch_base_02.st ---- *)
FUNCTION_BLOCK FB
VAR_INPUT
    runRequest      : BOOL;
    pressure        : REAL;
    pressureValid   : BOOL;
    fuelFlow        : REAL;
    steamFlow       : REAL;
    outletCmd       : INT;
    outletFeedback  : INT;
    resetBtn        : BOOL;
END_VAR
VAR_OUTPUT
    tripLatched     : BOOL;
    fuelPermit      : BOOL;
    currentCauseMask: WORD;
    latchedCauseMask: WORD;
    diagnosticActive: BOOL;
END_VAR
VAR
    prevResetBtn    : BOOL;
    valveStickingCnt: INT;
END_VAR
VAR_TEMP
    resetRising     : BOOL;
    tmpMask         : WORD;
    overpressure    : BOOL;
    valveCondition  : BOOL;
    combustionCond  : BOOL;
    unlocatedCond   : BOOL;
END_VAR
// ENGINEERING_CONTRACT
// PUB003: tripLatched activates on runRequest AND (NOT pressureValid OR pressure>=4500.0)
// PUB004: tripLatched holds until valid reset rising edge
// PUB005: reset requires resetBtn rising edge AND NOT runRequest AND pressureValid AND pressure<=4200.0
// PUB006: currentCauseMask low 4 bits: bit0=1 transmitter fail, bit1=2 valve sticking, bit2=4 combustion excess, bit3=8 unlocated
// PUB007: valve sticking requires 3 consecutive scans; any break (condition fail / pressure drop / invalid / stop) clears counter
// PUB010: 300kPa hysteresis (trip at 4500.0, reset at 4200.0)
// PUB012: latchedCauseMask accumulates via bitwise OR during tripLatched; only valid reset clears to 0
// PUB014: fuelPermit = runRequest AND NOT tripLatched
// PUB015: diagnosticActive = currentCauseMask <> 0
// PUB016: NOT runRequest forces currentCauseMask=0 (bits are mutually exclusive per N10-S15)
// PUB017-018: allowed mask values {0,1,2,4,6,8}; N10-S11 validates bit1 requires 3 consecutive scans
// PUB019-022: same-scan behavior - trip and currentCauseMask computed from current inputs each scan
// PUB023-026: latchedCauseMask is historical accumulator, not snapshot; preserves full trip footprint
(* CONTRACT_RULES [] *)
;

resetRising := resetBtn AND NOT prevResetBtn;

tmpMask := 0;
overpressure := runRequest AND pressureValid AND (pressure >= 4500.0);
unlocatedCond := FALSE;

IF NOT runRequest THEN
    currentCauseMask := 0;
    valveStickingCnt := 0;
    tmpMask := 0;
ELSIF NOT pressureValid THEN
    currentCauseMask := 1;  // bit0
    valveStickingCnt := 0;
    tmpMask := 0;
ELSE
    valveCondition := (outletCmd >= 50) AND (outletFeedback <= 10);
    IF overpressure AND valveCondition THEN
        valveStickingCnt := valveStickingCnt + 1;
    ELSE
        valveStickingCnt := 0;
    END_IF;

    combustionCond := (fuelFlow >= 4.0) AND (steamFlow <= 10.0);

    IF valveStickingCnt >= 3 THEN
        tmpMask := TO_WORD(TO_UINT(tmpMask) OR 2);  // bit1
    END_IF;

    IF combustionCond THEN
        tmpMask := TO_WORD(TO_UINT(tmpMask) OR 4);  // bit2
    END_IF;

    IF overpressure AND ((tmpMask AND 2) = 0) AND ((tmpMask AND 4) = 0) THEN
        tmpMask := TO_WORD(TO_UINT(tmpMask) OR 8);  // bit3 unlocated
    END_IF;

    currentCauseMask := tmpMask;
END_IF;

IF tripLatched THEN
    IF resetRising AND NOT runRequest AND pressureValid AND (pressure <= 4200.0) THEN
        tripLatched := FALSE;
        latchedCauseMask := 0;
    ELSE
        latchedCauseMask := TO_WORD(TO_UINT(latchedCauseMask) OR TO_UINT(currentCauseMask));
    END_IF;
ELSE
    IF runRequest AND (NOT pressureValid OR (pressure >= 4500.0)) THEN
        tripLatched := TRUE;
        latchedCauseMask := currentCauseMask;
    ELSE
        tripLatched := FALSE;
        latchedCauseMask := 0;
    END_IF;
END_IF;

fuelPermit := runRequest AND NOT tripLatched;

diagnosticActive := (currentCauseMask <> 0);

prevResetBtn := resetBtn;

END_FUNCTION_BLOCK

(* ---- self-hard-06.patch_base_03.st ---- *)
FUNCTION_BLOCK FB
VAR_INPUT
    runRequest      : BOOL;
    pressure        : REAL;
    pressureValid   : BOOL;
    fuelFlow        : REAL;
    steamFlow       : REAL;
    outletCmd       : INT;
    outletFeedback  : INT;
    resetBtn        : BOOL;
END_VAR
VAR_OUTPUT
    tripLatched     : BOOL;
    fuelPermit      : BOOL;
    currentCauseMask: WORD;
    latchedCauseMask: WORD;
    diagnosticActive: BOOL;
END_VAR
VAR
    prevResetBtn    : BOOL;
    valveStickingCnt: INT;
END_VAR
VAR_TEMP
    resetRising     : BOOL;
    tmpMask         : WORD;
    overpressure    : BOOL;
    valveCondition  : BOOL;
    combustionCond  : BOOL;
    unlocatedCond   : BOOL;
END_VAR
// ENGINEERING_CONTRACT
// PUB003: tripLatched activates on runRequest AND (NOT pressureValid OR pressure>=4500.0)
// PUB004: tripLatched holds until valid reset rising edge
// PUB005: reset requires resetBtn rising edge AND NOT runRequest AND pressureValid AND pressure<=4200.0
// PUB006: currentCauseMask low 4 bits: bit0=1 transmitter fail, bit1=2 valve sticking, bit2=4 combustion excess, bit3=8 unlocated
// PUB007: valve sticking requires 3 consecutive scans; any break (condition fail / pressure drop / invalid / stop) clears counter
// PUB010: 300kPa hysteresis (trip at 4500.0, reset at 4200.0)
// PUB012: latchedCauseMask accumulates via bitwise OR during tripLatched; only valid reset clears to 0
// PUB014: fuelPermit = runRequest AND NOT tripLatched
// PUB015: diagnosticActive = currentCauseMask <> 0
// PUB016: NOT runRequest forces currentCauseMask=0 (bits are mutually exclusive per N10-S15)
// PUB017-018: allowed mask values {0,1,2,4,6,8}; N10-S11 validates bit1 requires 3 consecutive scans
// PUB019-022: same-scan behavior - trip and currentCauseMask computed from current inputs each scan
// PUB023-026: latchedCauseMask is historical accumulator, not snapshot; preserves full trip footprint
(* CONTRACT_RULES [] *)
;

resetRising := resetBtn AND NOT prevResetBtn;

tmpMask := 0;
overpressure := runRequest AND pressureValid AND (pressure >= 4500.0);
unlocatedCond := FALSE;

IF NOT runRequest THEN
    currentCauseMask := 0;
    valveStickingCnt := 0;
    tmpMask := 0;
ELSIF NOT pressureValid THEN
    currentCauseMask := 1;  // bit0
    valveStickingCnt := 0;
    tmpMask := 0;
ELSE
    valveCondition := (outletCmd >= 50) AND (outletFeedback <= 10);
    IF overpressure AND valveCondition THEN
        valveStickingCnt := valveStickingCnt + 1;
    ELSE
        valveStickingCnt := 0;
    END_IF;

    combustionCond := (fuelFlow >= 4.0) AND (steamFlow <= 10.0);

    IF valveStickingCnt >= 3 THEN
        tmpMask := TO_WORD(TO_UINT(tmpMask) OR 2);  // bit1
    END_IF;

    IF combustionCond THEN
        tmpMask := TO_WORD(TO_UINT(tmpMask) OR 4);  // bit2
    END_IF;

    IF overpressure AND ((tmpMask AND 2) = 0) AND ((tmpMask AND 4) = 0) THEN
        tmpMask := TO_WORD(TO_UINT(tmpMask) OR 8);  // bit3 unlocated
    END_IF;

    currentCauseMask := tmpMask;
END_IF;

IF tripLatched THEN
    IF resetRising AND NOT runRequest AND pressureValid AND (pressure <= 4200.0) THEN
        tripLatched := FALSE;
        latchedCauseMask := 0;
    ELSE
        latchedCauseMask := TO_WORD(TO_UINT(latchedCauseMask) OR TO_UINT(currentCauseMask));
    END_IF;
ELSE
    IF runRequest AND (NOT pressureValid OR (pressure >= 4500.0)) THEN
        tripLatched := TRUE;
        latchedCauseMask := currentCauseMask;
    ELSE
        tripLatched := FALSE;
        latchedCauseMask := 0;
    END_IF;
END_IF;

fuelPermit := runRequest AND NOT tripLatched;

diagnosticActive := (currentCauseMask <> 0);

prevResetBtn := resetBtn;

END_FUNCTION_BLOCK

(* ---- self-hard-06.raw_candidate_01.st ---- *)
FUNCTION_BLOCK FB
VAR_INPUT
    runRequest      : BOOL;
    pressure        : REAL;
    pressureValid   : BOOL;
    fuelFlow        : REAL;
    steamFlow       : REAL;
    outletCmd       : INT;
    outletFeedback  : INT;
    resetBtn        : BOOL;
END_VAR
VAR_OUTPUT
    tripLatched     : BOOL;
    fuelPermit      : BOOL;
    currentCauseMask: WORD;
    latchedCauseMask: WORD;
    diagnosticActive: BOOL;
END_VAR
VAR
    prevResetBtn    : BOOL;
    valveStickingCnt: INT;
END_VAR
VAR_TEMP
    resetRising     : BOOL;
    tmpMask         : WORD;
    overpressure    : BOOL;
    valveCondition  : BOOL;
    combustionCond  : BOOL;
    unlocatedCond   : BOOL;
END_VAR
// ENGINEERING_CONTRACT
// PUB003: tripLatched activates on runRequest AND (NOT pressureValid OR pressure>=4500.0)
// PUB004: tripLatched holds until valid reset rising edge
// PUB005: reset requires resetBtn rising edge AND NOT runRequest AND pressureValid AND pressure<=4200.0
// PUB006: currentCauseMask low 4 bits: bit0=1 transmitter fail, bit1=2 valve sticking, bit2=4 combustion excess, bit3=8 unlocated
// PUB007: valve sticking requires 3 consecutive scans; any break (condition fail / pressure drop / invalid / stop) clears counter
// PUB010: 300kPa hysteresis (trip at 4500.0, reset at 4200.0)
// PUB012: latchedCauseMask accumulates via bitwise OR during tripLatched; only valid reset clears to 0
// PUB014: fuelPermit = runRequest AND NOT tripLatched
// PUB015: diagnosticActive = currentCauseMask <> 0
// PUB016: NOT runRequest forces currentCauseMask=0 (bits are mutually exclusive per N10-S15)
// PUB017-018: allowed mask values {0,1,2,4,6,8}; N10-S11 validates bit1 requires 3 consecutive scans
// PUB019-022: same-scan behavior - trip and currentCauseMask computed from current inputs each scan
// PUB023-026: latchedCauseMask is historical accumulator, not snapshot; preserves full trip footprint
(* CONTRACT_RULES [] *)
;

resetRising := resetBtn AND NOT prevResetBtn;

tmpMask := 0;
overpressure := runRequest AND pressureValid AND (pressure >= 4500.0);
unlocatedCond := FALSE;

IF NOT runRequest THEN
    currentCauseMask := 0;
    valveStickingCnt := 0;
    tmpMask := 0;
ELSIF NOT pressureValid THEN
    currentCauseMask := 1;  // bit0
    valveStickingCnt := 0;
    tmpMask := 0;
ELSE
    valveCondition := (outletCmd >= 50) AND (outletFeedback <= 10);
    IF overpressure AND valveCondition THEN
        valveStickingCnt := valveStickingCnt + 1;
    ELSE
        valveStickingCnt := 0;
    END_IF

    combustionCond := (fuelFlow >= 4.0) AND (steamFlow <= 10.0);

    IF valveStickingCnt >= 3 THEN
        tmpMask := TO_WORD(TO_UINT(tmpMask) OR 2);  // bit1
    END_IF;

    IF combustionCond THEN
        tmpMask := TO_WORD(TO_UINT(tmpMask) OR 4);  // bit2
    END_IF;

    IF overpressure AND ((tmpMask AND 2) = 0) AND ((tmpMask AND 4) = 0) THEN
        tmpMask := TO_WORD(TO_UINT(tmpMask) OR 8);  // bit3 unlocated
    END_IF;

    currentCauseMask := tmpMask;
END_IF;

IF tripLatched THEN
    IF resetRising AND NOT runRequest AND pressureValid AND (pressure <= 4200.0) THEN
        tripLatched := FALSE;
        latchedCauseMask := 0;
    ELSE
        latchedCauseMask := TO_WORD(TO_UINT(latchedCauseMask) OR TO_UINT(currentCauseMask));
    END_IF;
ELSE
    IF runRequest AND (NOT pressureValid OR (pressure >= 4500.0)) THEN
        tripLatched := TRUE;
        latchedCauseMask := currentCauseMask;
    ELSE
        tripLatched := FALSE;
        latchedCauseMask := 0;
    END_IF;
END_IF;

fuelPermit := runRequest AND NOT tripLatched;

diagnosticActive := (currentCauseMask <> 0);

prevResetBtn := resetBtn;

END_FUNCTION_BLOCK

(* ---- self-hard-07.candidate_01.st ---- *)
FUNCTION_BLOCK FB
VAR_INPUT
    mode            : INT;           (* 0=Manual 1=Auto 2=Cascade *)
    resetBtn        : BOOL;          (* Rising edge: reset to initial state *)
    scanSeconds     : REAL;          (* Scan period in seconds *)
    tempSP          : REAL;          (* Temperature setpoint, degC *)
    tempPV          : REAL;          (* Temperature process value, degC *)
    flowPV          : REAL;          (* Flow process value, t/h *)
    manualFlowSP    : REAL;          (* Manual flow setpoint, t/h *)
    manualValve     : REAL;          (* Manual valve position, % *)
END_VAR
VAR_OUTPUT
    flowSP          : REAL;          (* Flow setpoint output, t/h, clamped 0..50 *)
    valveCommand    : REAL;          (* Valve command output, %, clamped 0..100 *)
    fault           : BOOL;          (* Fault: invalid mode or scanSeconds *)
    normalMode      : BOOL;          (* This scan is normal operation (not reset/fault/switch/first) *)
END_VAR
VAR
    prevResetBtn    : BOOL    := FALSE;
    prevMode        : INT     := 0;
    accT            : REAL    := 0.0;    (* Integral state outer loop, unit t/h *)
    accF            : REAL    := 0.0;    (* Integral state inner loop, unit % *)
    firstScan       : BOOL    := TRUE;
END_VAR
VAR_TEMP
    tmpModeChanged  : BOOL;
    tmpET           : REAL;
    tmpEF           : REAL;
    tmpTrial        : REAL;
END_VAR
(*
ENGINEERING_CONTRACT:
  Modes: 0=Manual (both follow manual), 1=Auto (flow=manual, PI valve), 2=Cascade (PI flow then PI valve)
  Outputs: flowSP [0..50] t/h, valveCommand [0..100] %; retention per mode contract
  Activation: PI execution on normalMode=TRUE; bumpless transfer on mode switch (outputs hold/follow per spec)
  Reset/Deactivation: resetBtn rising edge → init to manual values, no PI on that scan
  Fault: mode∉{0,1,2} or scanSeconds∉(0,10] → fault, follow manual, no PI
  Priority: reset>fault (both reported), first-scan treated as switch (normalMode=FALSE)
  Units: KiT=0.2 (t/h)/(degC·s), KpT=1.0 (t/h)/degC; KiF=0.5 %/((t/h)·s), KpF=2.0 %/(t/h)
  Anti-windup: back-calculation from clamped output to accumulator
*)
BEGIN
    (* --- First scan: initialize outputs and accumulators --- *)
    IF firstScan THEN
        flowSP      := manualFlowSP;
        valveCommand := manualValve;
        accT        := 0.0;
        accF        := 0.0;
        fault       := FALSE;
        normalMode  := FALSE;
        firstScan   := FALSE;
        prevResetBtn := resetBtn;
        prevMode    := mode;
        RETURN;
    END_IF;

    (* --- Detect state changes --- *)
    tmpModeChanged := (mode <> prevMode);

    (* --- Reset rising edge: immediate fallback to manual, no PI this scan --- *)
    IF resetBtn AND NOT prevResetBtn THEN
        flowSP       := manualFlowSP;
        valveCommand := manualValve;
        accT         := 0.0;
        accF         := 0.0;
        fault        := FALSE;
        normalMode   := FALSE;
        prevResetBtn := resetBtn;
        prevMode     := mode;
        RETURN;
    END_IF;

    (* --- Fault condition: invalid mode or scanSeconds --- *)
    fault := (mode < 0) OR (mode > 2) OR (scanSeconds <= 0.0) OR (scanSeconds > 10.0);

    (* --- Fault fallback: follow manual immediately, no integral update --- *)
    IF fault THEN
        flowSP       := manualFlowSP;
        valveCommand := manualValve;
        accT         := 0.0;
        accF         := 0.0;
        normalMode   := FALSE;
        prevResetBtn := resetBtn;
        prevMode     := mode;
        RETURN;
    END_IF;

    (* --- Normal operation or mode-transition scan --- *)
    IF mode = 0 THEN
        (* Manual: both outputs follow manual values; recalc accumulators for bumpless re-entry *)
        flowSP       := manualFlowSP;
        valveCommand := manualValve;
        tmpET := tempSP - tempPV;
        tmpEF := flowSP - flowPV;
        accT := flowSP - 1.0 * tmpET;
        accF := valveCommand - 2.0 * tmpEF;

    ELSIF mode = 2 THEN
        (* Cascade: outer loop PI → flowSP; inner loop PI → valveCommand *)
        IF tmpModeChanged THEN
            (* Mode switch: hold outputs, recalc accumulators for bumpless transfer *)
            flowSP       := flowSP;
            valveCommand := valveCommand;
            tmpET := tempSP - tempPV;
            tmpEF := flowSP - flowPV;
            accT := flowSP - 1.0 * tmpET;
            accF := valveCommand - 2.0 * tmpEF;
        ELSE
            (* Normal PI execution with anti-windup back-calculation *)
            tmpET := tempSP - tempPV;
            tmpEF := flowSP - flowPV;
            (* Outer loop *)
            tmpTrial := accT + 0.2 * tmpET * scanSeconds;
            flowSP   := LIMIT(0.0, 1.0 * tmpET + tmpTrial, 50.0);
            accT     := flowSP - 1.0 * tmpET;
            (* Inner loop uses current flowSP *)
            tmpEF    := flowSP - flowPV;
            tmpTrial := accF + 0.5 * tmpEF * scanSeconds;
            valveCommand := LIMIT(0.0, 2.0 * tmpEF + tmpTrial, 100.0);
            accF     := valveCommand - 2.0 * tmpEF;
        END_IF;

    ELSIF mode = 1 THEN
        (* Auto: flowSP = manualFlowSP; inner loop PI → valveCommand *)
        IF tmpModeChanged THEN
            (* Mode switch: flowSP follows manual, valve holds; recalc accumulators *)
            flowSP       := manualFlowSP;
            valveCommand := valveCommand;
            tmpET := tempSP - tempPV;
            tmpEF := flowSP - flowPV;
            accT := flowSP - 1.0 * tmpET;
            accF := valveCommand - 2.0 * tmpEF;
        ELSE
            (* Normal PI execution *)
            flowSP       := manualFlowSP;
            tmpET        := tempSP - tempPV;
            accT         := flowSP - 1.0 * tmpET;
            tmpEF        := flowSP - flowPV;
            tmpTrial     := accF + 0.5 * tmpEF * scanSeconds;
            valveCommand := LIMIT(0.0, 2.0 * tmpEF + tmpTrial, 100.0);
            accF         := valveCommand - 2.0 * tmpEF;
        END_IF;
    END_IF;

    (* --- Update previous-state tracking --- *)
    prevResetBtn := resetBtn;
    prevMode     := mode;

    (* --- normalMode: second-or-later scan, stable mode, no fault, no reset rising edge --- *)
    normalMode := NOT firstScan AND (mode = prevMode) AND NOT fault AND NOT (resetBtn AND NOT prevResetBtn);
END_FUNCTION_BLOCK

(* ---- self-hard-07.patch_base_02.st ---- *)
FUNCTION_BLOCK FB
VAR_INPUT
    mode            : INT;           (* 0=Manual 1=Auto 2=Cascade *)
    resetBtn        : BOOL;          (* Rising edge: reset to initial state *)
    scanSeconds     : REAL;          (* Scan period in seconds *)
    tempSP          : REAL;          (* Temperature setpoint, degC *)
    tempPV          : REAL;          (* Temperature process value, degC *)
    flowPV          : REAL;          (* Flow process value, t/h *)
    manualFlowSP    : REAL;          (* Manual flow setpoint, t/h *)
    manualValve     : REAL;          (* Manual valve position, % *)
END_VAR
VAR_OUTPUT
    flowSP          : REAL;          (* Flow setpoint output, t/h, clamped 0..50 *)
    valveCommand    : REAL;          (* Valve command output, %, clamped 0..100 *)
    fault           : BOOL;          (* Fault: invalid mode or scanSeconds *)
    normalMode      : BOOL;          (* This scan is normal operation (not reset/fault/switch/first) *)
END_VAR
VAR
    prevResetBtn    : BOOL    := FALSE;
    prevMode        : INT     := 0;
    accT            : REAL    := 0.0;    (* Integral state outer loop, unit t/h *)
    accF            : REAL    := 0.0;    (* Integral state inner loop, unit % *)
    firstScan       : BOOL    := TRUE;
END_VAR
VAR_TEMP
    tmpModeChanged  : BOOL;
    tmpET           : REAL;
    tmpEF           : REAL;
    tmpTrial        : REAL;
END_VAR
(*
ENGINEERING_CONTRACT:
  Modes: 0=Manual (both follow manual), 1=Auto (flow=manual, PI valve), 2=Cascade (PI flow then PI valve)
  Outputs: flowSP [0..50] t/h, valveCommand [0..100] %; retention per mode contract
  Activation: PI execution on normalMode=TRUE; bumpless transfer on mode switch (outputs hold/follow per spec)
  Reset/Deactivation: resetBtn rising edge → init to manual values, no PI on that scan
  Fault: mode∉{0,1,2} or scanSeconds∉(0,10] → fault, follow manual, no PI
  Priority: reset>fault (both reported), first-scan treated as switch (normalMode=FALSE)
  Units: KiT=0.2 (t/h)/(degC·s), KpT=1.0 (t/h)/degC; KiF=0.5 %/((t/h)·s), KpF=2.0 %/(t/h)
  Anti-windup: back-calculation from clamped output to accumulator
*)
BEGIN
    (* --- First scan: initialize outputs and accumulators --- *)
    IF firstScan THEN
        flowSP      := manualFlowSP;
        valveCommand := manualValve;
        accT        := 0.0;
        accF        := 0.0;
        fault       := FALSE;
        normalMode  := FALSE;
        firstScan   := FALSE;
        prevResetBtn := resetBtn;
        prevMode    := mode;
        RETURN;
    END_IF;

    (* --- Detect state changes --- *)
    tmpModeChanged := (mode <> prevMode);

    (* --- Reset rising edge: immediate fallback to manual, no PI this scan --- *)
    IF resetBtn AND NOT prevResetBtn THEN
        flowSP       := manualFlowSP;
        valveCommand := manualValve;
        accT         := 0.0;
        accF         := 0.0;
        fault        := FALSE;
        normalMode   := FALSE;
        prevResetBtn := resetBtn;
        prevMode     := mode;
        RETURN;
    END_IF;

    (* --- Fault condition: invalid mode or scanSeconds --- *)
    fault := (mode < 0) OR (mode > 2) OR (scanSeconds <= 0.0) OR (scanSeconds > 10.0);

    (* --- Fault fallback: follow manual immediately, no integral update --- *)
    IF fault THEN
        flowSP       := manualFlowSP;
        valveCommand := manualValve;
        accT         := 0.0;
        accF         := 0.0;
        normalMode   := FALSE;
        prevResetBtn := resetBtn;
        prevMode     := mode;
        RETURN;
    END_IF;

    (* --- Normal operation or mode-transition scan --- *)
    IF mode = 0 THEN
        (* Manual: both outputs follow manual values; recalc accumulators for bumpless re-entry *)
        flowSP       := manualFlowSP;
        valveCommand := manualValve;
        tmpET := tempSP - tempPV;
        tmpEF := flowSP - flowPV;
        accT := flowSP - 1.0 * tmpET;
        accF := valveCommand - 2.0 * tmpEF;

    ELSIF mode = 2 THEN
        (* Cascade: outer loop PI → flowSP; inner loop PI → valveCommand *)
        IF tmpModeChanged THEN
            (* Mode switch: hold outputs, recalc accumulators for bumpless transfer *)
            flowSP       := flowSP;
            valveCommand := valveCommand;
            tmpET := tempSP - tempPV;
            tmpEF := flowSP - flowPV;
            accT := flowSP - 1.0 * tmpET;
            accF := valveCommand - 2.0 * tmpEF;
        ELSE
            (* Normal PI execution with anti-windup back-calculation *)
            tmpET := tempSP - tempPV;
            tmpEF := flowSP - flowPV;
            (* Outer loop *)
            tmpTrial := accT + 0.2 * tmpET * scanSeconds;
            flowSP   := LIMIT(0.0, 1.0 * tmpET + tmpTrial, 50.0);
            accT     := flowSP - 1.0 * tmpET;
            (* Inner loop uses current flowSP *)
            tmpEF    := flowSP - flowPV;
            tmpTrial := accF + 0.5 * tmpEF * scanSeconds;
            valveCommand := LIMIT(0.0, 2.0 * tmpEF + tmpTrial, 100.0);
            accF     := valveCommand - 2.0 * tmpEF;
        END_IF;

    ELSIF mode = 1 THEN
        (* Auto: flowSP = manualFlowSP; inner loop PI → valveCommand *)
        IF tmpModeChanged THEN
            (* Mode switch: flowSP follows manual, valve holds; recalc accumulators *)
            flowSP       := manualFlowSP;
            valveCommand := valveCommand;
            tmpET := tempSP - tempPV;
            tmpEF := flowSP - flowPV;
            accT := flowSP - 1.0 * tmpET;
            accF := valveCommand - 2.0 * tmpEF;
        ELSE
            (* Normal PI execution *)
            flowSP       := manualFlowSP;
            tmpET        := tempSP - tempPV;
            accT         := flowSP - 1.0 * tmpET;
            tmpEF        := flowSP - flowPV;
            tmpTrial     := accF + 0.5 * tmpEF * scanSeconds;
            valveCommand := LIMIT(0.0, 2.0 * tmpEF + tmpTrial, 100.0);
            accF         := valveCommand - 2.0 * tmpEF;
        END_IF;
    END_IF;

    (* --- Update previous-state tracking --- *)
    prevResetBtn := resetBtn;
    prevMode     := mode;

    (* --- normalMode: second-or-later scan, stable mode, no fault, no reset rising edge --- *)
    normalMode := NOT firstScan AND (mode = prevMode) AND NOT fault AND NOT (resetBtn AND NOT prevResetBtn);
END_FUNCTION_BLOCK

(* ---- self-hard-07.patch_base_03.st ---- *)
FUNCTION_BLOCK FB
VAR_INPUT
    mode            : INT;           (* 0=Manual 1=Auto 2=Cascade *)
    resetBtn        : BOOL;          (* Rising edge: reset to initial state *)
    scanSeconds     : REAL;          (* Scan period in seconds *)
    tempSP          : REAL;          (* Temperature setpoint, degC *)
    tempPV          : REAL;          (* Temperature process value, degC *)
    flowPV          : REAL;          (* Flow process value, t/h *)
    manualFlowSP    : REAL;          (* Manual flow setpoint, t/h *)
    manualValve     : REAL;          (* Manual valve position, % *)
END_VAR
VAR_OUTPUT
    flowSP          : REAL;          (* Flow setpoint output, t/h, clamped 0..50 *)
    valveCommand    : REAL;          (* Valve command output, %, clamped 0..100 *)
    fault           : BOOL;          (* Fault: invalid mode or scanSeconds *)
    normalMode      : BOOL;          (* This scan is normal operation (not reset/fault/switch/first) *)
END_VAR
VAR
    prevResetBtn    : BOOL    := FALSE;
    prevMode        : INT     := 0;
    accT            : REAL    := 0.0;    (* Integral state outer loop, unit t/h *)
    accF            : REAL    := 0.0;    (* Integral state inner loop, unit % *)
    firstScan       : BOOL    := TRUE;
END_VAR
VAR_TEMP
    tmpModeChanged  : BOOL;
    tmpET           : REAL;
    tmpEF           : REAL;
    tmpTrial        : REAL;
END_VAR
(*
ENGINEERING_CONTRACT:
  Modes: 0=Manual (both follow manual), 1=Auto (flow=manual, PI valve), 2=Cascade (PI flow then PI valve)
  Outputs: flowSP [0..50] t/h, valveCommand [0..100] %; retention per mode contract
  Activation: PI execution on normalMode=TRUE; bumpless transfer on mode switch (outputs hold/follow per spec)
  Reset/Deactivation: resetBtn rising edge → init to manual values, no PI on that scan
  Fault: mode∉{0,1,2} or scanSeconds∉(0,10] → fault, follow manual, no PI
  Priority: reset>fault (both reported), first-scan treated as switch (normalMode=FALSE)
  Units: KiT=0.2 (t/h)/(degC·s), KpT=1.0 (t/h)/degC; KiF=0.5 %/((t/h)·s), KpF=2.0 %/(t/h)
  Anti-windup: back-calculation from clamped output to accumulator
*)
BEGIN
    (* --- First scan: initialize outputs and accumulators --- *)
    IF firstScan THEN
        flowSP      := manualFlowSP;
        valveCommand := manualValve;
        accT        := 0.0;
        accF        := 0.0;
        fault       := FALSE;
        normalMode  := FALSE;
        firstScan   := FALSE;
        prevResetBtn := resetBtn;
        prevMode    := mode;
        RETURN;
    END_IF;

    (* --- Detect state changes --- *)
    tmpModeChanged := (mode <> prevMode);

    (* --- Reset rising edge: immediate fallback to manual, no PI this scan --- *)
    IF resetBtn AND NOT prevResetBtn THEN
        flowSP       := manualFlowSP;
        valveCommand := manualValve;
        accT         := 0.0;
        accF         := 0.0;
        fault        := FALSE;
        normalMode   := FALSE;
        prevResetBtn := resetBtn;
        prevMode     := mode;
        RETURN;
    END_IF;

    (* --- Fault condition: invalid mode or scanSeconds --- *)
    fault := (mode < 0) OR (mode > 2) OR (scanSeconds <= 0.0) OR (scanSeconds > 10.0);

    (* --- Fault fallback: follow manual immediately, no integral update --- *)
    IF fault THEN
        flowSP       := manualFlowSP;
        valveCommand := manualValve;
        accT         := 0.0;
        accF         := 0.0;
        normalMode   := FALSE;
        prevResetBtn := resetBtn;
        prevMode     := mode;
        RETURN;
    END_IF;

    (* --- Normal operation or mode-transition scan --- *)
    IF mode = 0 THEN
        (* Manual: both outputs follow manual values; recalc accumulators for bumpless re-entry *)
        flowSP       := manualFlowSP;
        valveCommand := manualValve;
        tmpET := tempSP - tempPV;
        tmpEF := flowSP - flowPV;
        accT := flowSP - 1.0 * tmpET;
        accF := valveCommand - 2.0 * tmpEF;

    ELSIF mode = 2 THEN
        (* Cascade: outer loop PI → flowSP; inner loop PI → valveCommand *)
        IF tmpModeChanged THEN
            (* Mode switch: hold outputs, recalc accumulators for bumpless transfer *)
            flowSP       := flowSP;
            valveCommand := valveCommand;
            tmpET := tempSP - tempPV;
            tmpEF := flowSP - flowPV;
            accT := flowSP - 1.0 * tmpET;
            accF := valveCommand - 2.0 * tmpEF;
        ELSE
            (* Normal PI execution with anti-windup back-calculation *)
            tmpET := tempSP - tempPV;
            tmpEF := flowSP - flowPV;
            (* Outer loop *)
            tmpTrial := accT + 0.2 * tmpET * scanSeconds;
            flowSP   := LIMIT(0.0, 1.0 * tmpET + tmpTrial, 50.0);
            accT     := flowSP - 1.0 * tmpET;
            (* Inner loop uses current flowSP *)
            tmpEF    := flowSP - flowPV;
            tmpTrial := accF + 0.5 * tmpEF * scanSeconds;
            valveCommand := LIMIT(0.0, 2.0 * tmpEF + tmpTrial, 100.0);
            accF     := valveCommand - 2.0 * tmpEF;
        END_IF;

    ELSIF mode = 1 THEN
        (* Auto: flowSP = manualFlowSP; inner loop PI → valveCommand *)
        IF tmpModeChanged THEN
            (* Mode switch: flowSP follows manual, valve holds; recalc accumulators *)
            flowSP       := manualFlowSP;
            valveCommand := valveCommand;
            tmpET := tempSP - tempPV;
            tmpEF := flowSP - flowPV;
            accT := flowSP - 1.0 * tmpET;
            accF := valveCommand - 2.0 * tmpEF;
        ELSE
            (* Normal PI execution *)
            flowSP       := manualFlowSP;
            tmpET        := tempSP - tempPV;
            accT         := flowSP - 1.0 * tmpET;
            tmpEF        := flowSP - flowPV;
            tmpTrial     := accF + 0.5 * tmpEF * scanSeconds;
            valveCommand := LIMIT(0.0, 2.0 * tmpEF + tmpTrial, 100.0);
            accF         := valveCommand - 2.0 * tmpEF;
        END_IF;
    END_IF;

    (* --- Update previous-state tracking --- *)
    prevResetBtn := resetBtn;
    prevMode     := mode;

    (* --- normalMode: second-or-later scan, stable mode, no fault, no reset rising edge --- *)
    normalMode := NOT firstScan AND (mode = prevMode) AND NOT fault AND NOT (resetBtn AND NOT prevResetBtn);
END_FUNCTION_BLOCK

(* ---- self-hard-07.raw_candidate_01.st ---- *)
FUNCTION_BLOCK FB
VAR_INPUT
    mode            : INT;           (* 0=Manual 1=Auto 2=Cascade *)
    resetBtn        : BOOL;          (* Rising edge: reset to initial state *)
    scanSeconds     : REAL;          (* Scan period in seconds *)
    tempSP          : REAL;          (* Temperature setpoint, degC *)
    tempPV          : REAL;          (* Temperature process value, degC *)
    flowPV          : REAL;          (* Flow process value, t/h *)
    manualFlowSP    : REAL;          (* Manual flow setpoint, t/h *)
    manualValve     : REAL;          (* Manual valve position, % *)
END_VAR
VAR_OUTPUT
    flowSP          : REAL;          (* Flow setpoint output, t/h, clamped 0..50 *)
    valveCommand    : REAL;          (* Valve command output, %, clamped 0..100 *)
    fault           : BOOL;          (* Fault: invalid mode or scanSeconds *)
    normalMode      : BOOL;          (* This scan is normal operation (not reset/fault/switch/first) *)
END_VAR
VAR
    prevResetBtn    : BOOL    := FALSE;
    prevMode        : INT     := 0;
    accT            : REAL    := 0.0;    (* Integral state outer loop, unit t/h *)
    accF            : REAL    := 0.0;    (* Integral state inner loop, unit % *)
    firstScan       : BOOL    := TRUE;
END_VAR
VAR_TEMP
    tmpModeChanged  : BOOL;
    tmpET           : REAL;
    tmpEF           : REAL;
    tmpTrial        : REAL;
END_VAR
(*
ENGINEERING_CONTRACT:
  Modes: 0=Manual (both follow manual), 1=Auto (flow=manual, PI valve), 2=Cascade (PI flow then PI valve)
  Outputs: flowSP [0..50] t/h, valveCommand [0..100] %; retention per mode contract
  Activation: PI execution on normalMode=TRUE; bumpless transfer on mode switch (outputs hold/follow per spec)
  Reset/Deactivation: resetBtn rising edge → init to manual values, no PI on that scan
  Fault: mode∉{0,1,2} or scanSeconds∉(0,10] → fault, follow manual, no PI
  Priority: reset>fault (both reported), first-scan treated as switch (normalMode=FALSE)
  Units: KiT=0.2 (t/h)/(degC·s), KpT=1.0 (t/h)/degC; KiF=0.5 %/((t/h)·s), KpF=2.0 %/(t/h)
  Anti-windup: back-calculation from clamped output to accumulator
*)
BEGIN
    (* --- First scan: initialize outputs and accumulators --- *)
    IF firstScan THEN
        flowSP      := manualFlowSP;
        valveCommand := manualValve;
        accT        := 0.0;
        accF        := 0.0;
        fault       := FALSE;
        normalMode  := FALSE;
        firstScan   := FALSE;
        prevResetBtn := resetBtn;
        prevMode    := mode;
        RETURN;
    END_IF

    (* --- Detect state changes --- *)
    tmpModeChanged := (mode <> prevMode);

    (* --- Reset rising edge: immediate fallback to manual, no PI this scan --- *)
    IF resetBtn AND NOT prevResetBtn THEN
        flowSP       := manualFlowSP;
        valveCommand := manualValve;
        accT         := 0.0;
        accF         := 0.0;
        fault        := FALSE;
        normalMode   := FALSE;
        prevResetBtn := resetBtn;
        prevMode     := mode;
        RETURN;
    END_IF

    (* --- Fault condition: invalid mode or scanSeconds --- *)
    fault := (mode < 0) OR (mode > 2) OR (scanSeconds <= 0.0) OR (scanSeconds > 10.0);

    (* --- Fault fallback: follow manual immediately, no integral update --- *)
    IF fault THEN
        flowSP       := manualFlowSP;
        valveCommand := manualValve;
        accT         := 0.0;
        accF         := 0.0;
        normalMode   := FALSE;
        prevResetBtn := resetBtn;
        prevMode     := mode;
        RETURN;
    END_IF

    (* --- Normal operation or mode-transition scan --- *)
    IF mode = 0 THEN
        (* Manual: both outputs follow manual values; recalc accumulators for bumpless re-entry *)
        flowSP       := manualFlowSP;
        valveCommand := manualValve;
        tmpET := tempSP - tempPV;
        tmpEF := flowSP - flowPV;
        accT := flowSP - 1.0 * tmpET;
        accF := valveCommand - 2.0 * tmpEF;

    ELSIF mode = 2 THEN
        (* Cascade: outer loop PI → flowSP; inner loop PI → valveCommand *)
        IF tmpModeChanged THEN
            (* Mode switch: hold outputs, recalc accumulators for bumpless transfer *)
            flowSP       := flowSP;
            valveCommand := valveCommand;
            tmpET := tempSP - tempPV;
            tmpEF := flowSP - flowPV;
            accT := flowSP - 1.0 * tmpET;
            accF := valveCommand - 2.0 * tmpEF;
        ELSE
            (* Normal PI execution with anti-windup back-calculation *)
            tmpET := tempSP - tempPV;
            tmpEF := flowSP - flowPV;
            (* Outer loop *)
            tmpTrial := accT + 0.2 * tmpET * scanSeconds;
            flowSP   := LIMIT(0.0, 1.0 * tmpET + tmpTrial, 50.0);
            accT     := flowSP - 1.0 * tmpET;
            (* Inner loop uses current flowSP *)
            tmpEF    := flowSP - flowPV;
            tmpTrial := accF + 0.5 * tmpEF * scanSeconds;
            valveCommand := LIMIT(0.0, 2.0 * tmpEF + tmpTrial, 100.0);
            accF     := valveCommand - 2.0 * tmpEF;
        END_IF

    ELSIF mode = 1 THEN
        (* Auto: flowSP = manualFlowSP; inner loop PI → valveCommand *)
        IF tmpModeChanged THEN
            (* Mode switch: flowSP follows manual, valve holds; recalc accumulators *)
            flowSP       := manualFlowSP;
            valveCommand := valveCommand;
            tmpET := tempSP - tempPV;
            tmpEF := flowSP - flowPV;
            accT := flowSP - 1.0 * tmpET;
            accF := valveCommand - 2.0 * tmpEF;
        ELSE
            (* Normal PI execution *)
            flowSP       := manualFlowSP;
            tmpET        := tempSP - tempPV;
            accT         := flowSP - 1.0 * tmpET;
            tmpEF        := flowSP - flowPV;
            tmpTrial     := accF + 0.5 * tmpEF * scanSeconds;
            valveCommand := LIMIT(0.0, 2.0 * tmpEF + tmpTrial, 100.0);
            accF         := valveCommand - 2.0 * tmpEF;
        END_IF;
    END_IF;

    (* --- Update previous-state tracking --- *)
    prevResetBtn := resetBtn;
    prevMode     := mode;

    (* --- normalMode: second-or-later scan, stable mode, no fault, no reset rising edge --- *)
    normalMode := NOT firstScan AND (mode = prevMode) AND NOT fault AND NOT (resetBtn AND NOT prevResetBtn);
END_FUNCTION_BLOCK
